      R_f[3,4] := -0.85727531;
      R_f[3,5] := 0.70266402;
      R_f[3,6] := -0.55573398;
      R_f[3,7] := 0.45469028;
      R_f[3,8] := -0.39782384;
      R_f[3,9] := 0.23143867;
      R_f[3,10] := -0.86177999;
      R_f[3,11] := 0.29983264;
      R_f[3,12] := 1.36218679;
      R_f[3,13] := 0.10939779;
      R_f[3,14] := -0.13315666;
      R_f[3,15] := -1.31117058;
      R_f[3,16] := 0.66998744;
      R_f[3,17] := 1.24320877;
      R_f[3,18] := -0.37031132;
      R_f[3,19] := -0.39300495;
      R_f[3,20] := -0.30342990;
      R_f[3,21] := -0.45216727;
      R_f[3,22] := -0.51143724;
      R_f[3,23] := 0.47799069;
      R_f[3,24] := -0.01827676;
      R_f[3,25] := 0.02519570;
      R_f[3,26] := 0.18636933;
      R_f[3,27] := -0.93594962;
      R_f[3,28] := 0.64644384;
      R_f[3,29] := -0.69783551;
      R_f[3,30] := -0.03558157;
      R_f[3,31] := 0.26994738;
      R_f[4,0] := -0.39344388;
      R_f[4,1] := 0.36222264;
      R_f[4,2] := -0.42310888;
      R_f[4,3] := 0.14989485;
      R_f[4,4] := -0.99088651;
      R_f[4,5] := 0.05782998;
      R_f[4,6] := 0.12812723;
      R_f[4,7] := -0.16467652;
      R_f[4,8] := -0.34736815;
      R_f[4,9] := 0.14911307;
      R_f[4,10] := 0.64495277;
      R_f[4,11] := 0.13966881;
      R_f[4,12] := 0.29640356;
      R_f[4,13] := 0.48785415;
      R_f[4,14] := -0.23574533;
      R_f[4,15] := 0.47339493;
      R_f[4,16] := -0.38768038;
      R_f[4,17] := 0.06993198;
      R_f[4,18] := 1.34699011;
      R_f[4,19] := -0.45494819;
      R_f[4,20] := -1.02421069;
      R_f[4,21] := 0.39080855;
      R_f[4,22] := -0.25200650;
      R_f[4,23] := 0.10465910;
      R_f[4,24] := 0.27367991;
      R_f[4,25] := 0.45886528;
      R_f[4,26] := 0.23802078;
      R_f[4,27] := -0.31698900;
      R_f[4,28] := 0.36807117;
      R_f[4,29] := -0.10262590;
      R_f[4,30] := -0.79831642;
      R_f[4,31] := 0.12268136;
      R_f[5,0] := 0.09268615;
      R_f[5,1] := 0.21935971;
      R_f[5,2] := -0.28605691;
      R_f[5,3] := -0.35209230;
      R_f[5,4] := 0.60323030;
      R_f[5,5] := -1.86963761;
      R_f[5,6] := 0.17267105;
      R_f[5,7] := 0.31667727;
      R_f[5,8] := 1.22614503;
      R_f[5,9] := -0.31814456;
      R_f[5,10] := 0.28639799;
      R_f[5,11] := 0.45808375;
      R_f[5,12] := 0.16454318;
      R_f[5,13] := -0.37628773;
      R_f[5,14] := 0.11079943;
      R_f[5,15] := 0.43248567;
      R_f[5,16] := 0.62867469;
      R_f[5,17] := -0.18534793;
      R_f[5,18] := -0.21310599;
      R_f[5,19] := -0.12530403;
      R_f[5,20] := -0.11672303;
      R_f[5,21] := -0.34058103;
      R_f[5,22] := 0.53213966;
      R_f[5,23] := -0.06069790;
      R_f[5,24] := 1.12480652;
      R_f[5,25] := -0.11877894;
      R_f[5,26] := 0.34038293;
      R_f[5,27] := 0.99329889;
      R_f[5,28] := 0.00048804;
      R_f[5,29] := -0.15688728;
      R_f[5,30] := 0.46641046;
      R_f[5,31] := 1.20925903;
      R_f[6,0] := -0.20363854;
      R_f[6,1] := -0.32236105;
      R_f[6,2] := -0.30276120;
      R_f[6,3] := -0.07836054;
      R_f[6,4] := 0.90966666;
      R_f[6,5] := 0.01400341;
      R_f[6,6] := 0.27368066;
      R_f[6,7] := 1.16410792;
      R_f[6,8] := 0.91342974;
      R_f[6,9] := -0.62499738;
      R_f[6,10] := 0.21230549;
      R_f[6,11] := 0.48843908;
      R_f[6,12] := -0.04002659;
      R_f[6,13] := -0.89160722;
      R_f[6,14] := 0.44720122;
      R_f[6,15] := -0.37033880;
      R_f[6,16] := 0.36007941;
      R_f[6,17] := 0.49022290;
      R_f[6,18] := -0.63365066;
      R_f[6,19] := -0.44222319;
      R_f[6,20] := 0.07470856;
      R_f[6,21] := -0.18424936;
      R_f[6,22] := -1.06331885;
      R_f[6,23] := 0.11231405;
      R_f[6,24] := 0.48846784;
      R_f[6,25] := 0.32240003;
      R_f[6,26] := -0.02514423;
      R_f[6,27] := 0.52824306;
      R_f[6,28] := 0.10916118;
      R_f[6,29] := 1.10423243;
      R_f[6,30] := 0.87132770;
      R_f[6,31] := -0.22497243;
      R_f[7,0] := 0.00290798;
      R_f[7,1] := 0.02380353;
      R_f[7,2] := -0.43460667;
      R_f[7,3] := -0.61469567;
      R_f[7,4] := 0.93173164;
      R_f[7,5] := -0.90107012;
      R_f[7,6] := 0.16509961;
      R_f[7,7] := 2.32758498;
      R_f[7,8] := -0.52484536;
      R_f[7,9] := 0.39195865;
      R_f[7,10] := -0.23609044;
      R_f[7,11] := 0.05608457;
      R_f[7,12] := -0.42776030;
      R_f[7,13] := -0.10564836;
      R_f[7,14] := -0.42611927;
      R_f[7,15] := -0.13254717;
      R_f[7,16] := 0.84613299;
      R_f[7,17] := -0.23140904;
      R_f[7,18] := 0.90073472;
      R_f[7,19] := -0.36597919;
      R_f[7,20] := 0.47446036;
      R_f[7,21] := -0.08705632;
      R_f[7,22] := -1.52176034;
      R_f[7,23] := 0.22270711;
      R_f[7,24] := -0.03422754;
      R_f[7,25] := 0.07659206;
      R_f[7,26] := 0.36599547;
      R_f[7,27] := -0.52767622;
      R_f[7,28] := -0.06631206;
      R_f[7,29] := -0.18978609;
      R_f[7,30] := 0.17292330;
      R_f[7,31] := 0.92969888;
      R_f[8,0] := -0.30634153;
      R_f[8,1] := -0.81952202;
      R_f[8,2] := -0.03526760;
      R_f[8,3] := -1.29526353;
      R_f[8,4] := 0.32094973;
      R_f[8,5] := -1.85603750;
      R_f[8,6] := 0.28356239;
      R_f[8,7] := 0.57538003;
      R_f[8,8] := -0.11039671;
      R_f[8,9] := -2.10963488;
      R_f[8,10] := -1.19219816;
      R_f[8,11] := -0.79363817;
      R_f[8,12] := 0.48992485;
      R_f[8,13] := 0.30308276;
      R_f[8,14] := 0.04908920;
      R_f[8,15] := 0.13945648;
      R_f[8,16] := -1.37335110;
      R_f[8,17] := 0.59385890;
      R_f[8,18] := -1.01455212;
      R_f[8,19] := -1.58437848;
      R_f[8,20] := -0.19760673;
      R_f[8,21] := -0.34158847;
      R_f[8,22] := 1.34096205;
      R_f[8,23] := 0.40719572;
      R_f[8,24] := -0.24326721;
      R_f[8,25] := -1.13661909;
      R_f[8,26] := -0.63606089;
      R_f[8,27] := 0.39769849;
      R_f[8,28] := -1.44548726;
      R_f[8,29] := 0.17782873;
      R_f[8,30] := -0.33304986;
      R_f[8,31] := -0.34794864;
      R_f[9,0] := -0.44309428;
      R_f[9,1] := -0.30440933;
      R_f[9,2] := 0.24199238;
      R_f[9,3] := 0.21034531;
      R_f[9,4] := -0.17321667;
      R_f[9,5] := -0.30677229;
      R_f[9,6] := -0.13734587;
      R_f[9,7] := 0.34537369;
      R_f[9,8] := -0.26872745;
      R_f[9,9] := 1.84128654;
      R_f[9,10] := 0.52121741;
      R_f[9,11] := 0.30513665;
      R_f[9,12] := -0.01998700;
      R_f[9,13] := -0.72075009;
      R_f[9,14] := -0.55062896;
      R_f[9,15] := -0.11161942;
      R_f[9,16] := 0.10928833;
      R_f[9,17] := 0.69333780;
      R_f[9,18] := -0.61185640;
      R_f[9,19] := -0.22928748;
      R_f[9,20] := 0.53006452;
      R_f[9,21] := 0.10420142;
      R_f[9,22] := -0.16613784;
      R_f[9,23] := 0.12584257;
      R_f[9,24] := 0.24575511;
      R_f[9,25] := 0.07394662;
      R_f[9,26] := 0.62375677;
      R_f[9,27] := 0.53293931;
      R_f[9,28] := 0.20416169;
      R_f[9,29] := -0.02031298;
      R_f[9,30] := -0.10528360;
      R_f[9,31] := 0.45511815;
      R_f[10,0] := 0.83232188;
      R_f[10,1] := -0.08258834;
      R_f[10,2] := -0.06935453;
      R_f[10,3] := 0.07768326;
      R_f[10,4] := 0.24524604;
      R_f[10,5] := -0.22525373;
      R_f[10,6] := 0.40935123;
      R_f[10,7] := -0.17911816;
      R_f[10,8] := -0.32271239;
      R_f[10,9] := -0.36832979;
      R_f[10,10] := -2.49958277;
      R_f[10,11] := -0.03748730;
      R_f[10,12] := -0.07992049;
      R_f[10,13] := 0.08578819;
      R_f[10,14] := -0.19220759;
      R_f[10,15] := 0.08966637;
      R_f[10,16] := -0.39432195;
      R_f[10,17] := 0.22714733;
      R_f[10,18] := -0.43346864;
      R_f[10,19] := -0.11305624;
      R_f[10,20] := 0.16338432;
      R_f[10,21] := -0.10953200;
      R_f[10,22] := -0.13001373;
      R_f[10,23] := 0.22707058;
      R_f[10,24] := 0.41991970;
      R_f[10,25] := 0.43455145;
      R_f[10,26] := 0.19583054;
      R_f[10,27] := 0.56395984;
      R_f[10,28] := -0.48473257;
      R_f[10,29] := 0.18865864;
      R_f[10,30] := 0.19654989;
      R_f[10,31] := 0.09913722;
      R_f[11,0] := 0.42754596;
      R_f[11,1] := 0.09423707;
      R_f[11,2] := -0.29017773;
      R_f[11,3] := -0.11189838;
      R_f[11,4] := -0.21009797;
      R_f[11,5] := -0.48191920;
      R_f[11,6] := 0.12651034;
      R_f[11,7] := 0.05790544;
      R_f[11,8] := -0.12319141;
      R_f[11,9] := 0.39675516;
      R_f[11,10] := -0.16217400;
      R_f[11,11] := 0.18192010;
      R_f[11,12] := 0.14949840;
      R_f[11,13] := -0.03762484;
      R_f[11,14] := -0.68928587;
      R_f[11,15] := 0.11334433;
      R_f[11,16] := -0.28812110;
      R_f[11,17] := 0.10144100;
      R_f[11,18] := -0.44992569;
      R_f[11,19] := -0.15579885;
      R_f[11,20] := -0.29591924;
      R_f[11,21] := -0.15366313;
      R_f[11,22] := -0.01909444;
      R_f[11,23] := 0.04565328;
      R_f[11,24] := -0.30796039;
      R_f[11,25] := -0.08308777;
      R_f[11,26] := 0.22044559;
      R_f[11,27] := 0.10441495;
      R_f[11,28] := 0.06342443;
      R_f[11,29] := -0.48254472;
      R_f[11,30] := 0.09183690;
      R_f[11,31] := -0.09384891;
      R_f[12,0] := 0.47012070;
      R_f[12,1] := -0.33459604;
      R_f[12,2] := -0.69821233;
      R_f[12,3] := 0.03733517;
      R_f[12,4] := 1.01428008;
      R_f[12,5] := -1.34689188;
      R_f[12,6] := 0.60434407;
      R_f[12,7] := 1.02553523;
      R_f[12,8] := 0.34444749;
      R_f[12,9] := -0.69957334;
      R_f[12,10] := 0.80366671;
      R_f[12,11] := 0.17610356;
      R_f[12,12] := 0.55641246;
      R_f[12,13] := -0.21217743;
      R_f[12,14] := -0.63918966;
      R_f[12,15] := -0.16232961;
      R_f[12,16] := 0.68742597;
      R_f[12,17] := 0.52715355;
      R_f[12,18] := 0.04790421;
      R_f[12,19] := -0.58621752;
      R_f[12,20] := 0.26796517;
      R_f[12,21] := -0.04791349;
      R_f[12,22] := -0.09341484;
      R_f[12,23] := 0.66781473;
      R_f[12,24] := 0.52626812;
      R_f[12,25] := 0.37837932;
      R_f[12,26] := 0.38251483;
      R_f[12,27] := 0.31467408;
      R_f[12,28] := -0.29517949;
      R_f[12,29] := -0.02343472;
      R_f[12,30] := 0.19953103;
      R_f[12,31] := 0.04299867;
      R_f[13,0] := 0.08943395;
      R_f[13,1] := -0.41928035;
      R_f[13,2] := -0.46420595;
      R_f[13,3] := -0.93849921;
      R_f[13,4] := 1.81882250;
      R_f[13,5] := -0.04638388;
      R_f[13,6] := -0.10525256;
      R_f[13,7] := -0.14901699;
      R_f[13,8] := 1.56855416;
      R_f[13,9] := -1.47332811;
      R_f[13,10] := 1.70304513;
      R_f[13,11] := 0.27727890;
      R_f[13,12] := 0.29618439;
      R_f[13,13] := 0.20549068;
      R_f[13,14] := 0.08464767;
      R_f[13,15] := -0.28658184;
      R_f[13,16] := 0.52141178;
      R_f[13,17] := -0.45672634;
      R_f[13,18] := -1.07117772;
      R_f[13,19] := -0.12635788;
      R_f[13,20] := -0.17076187;
      R_f[13,21] := -0.39133579;
      R_f[13,22] := -1.30128396;
      R_f[13,23] := -0.51295263;
      R_f[13,24] := 0.59420377;
      R_f[13,25] := -0.22949216;
      R_f[13,26] := -0.07507192;
      R_f[13,27] := 0.62209141;
      R_f[13,28] := -0.39097649;
      R_f[13,29] := 0.46184129;
      R_f[13,30] := 0.24478418;
      R_f[13,31] := 1.16894412;
      R_f[14,0] := 0.05281359;
      R_f[14,1] := -0.53310943;
      R_f[14,2] := -0.93560243;
      R_f[14,3] := 0.24883044;
      R_f[14,4] := -0.87425369;
      R_f[14,5] := 0.40351281;
      R_f[14,6] := -0.38772595;
      R_f[14,7] := 0.02093324;
      R_f[14,8] := -0.35284448;
      R_f[14,9] := -0.49149925;
      R_f[14,10] := 0.40103057;
      R_f[14,11] := -0.23631869;
      R_f[14,12] := -0.18181595;
      R_f[14,13] := 1.02885425;
      R_f[14,14] := 1.01850176;
      R_f[14,15] := 0.01374859;
      R_f[14,16] := 0.09904287;
      R_f[14,17] := 0.39969888;
      R_f[14,18] := 0.29445514;
      R_f[14,19] := -0.66422909;
      R_f[14,20] := 0.56930321;
      R_f[14,21] := 0.16506715;
      R_f[14,22] := -0.23321085;
      R_f[14,23] := 0.48102799;
      R_f[14,24] := -0.53297859;
      R_f[14,25] := 0.40016001;
      R_f[14,26] := -0.33044472;
      R_f[14,27] := 0.31068552;
      R_f[14,28] := 0.16014290;
      R_f[14,29] := 0.17083554;
      R_f[14,30] := 0.17105293;
      R_f[14,31] := 0.35666907;
      R_f[15,0] := 0.06514452;
      R_f[15,1] := -0.19740443;
      R_f[15,2] := 0.02617185;
      R_f[15,3] := 0.07652328;
      R_f[15,4] := 0.38803399;
      R_f[15,5] := -0.20535301;
      R_f[15,6] := -0.18448971;
      R_f[15,7] := -0.05007682;
      R_f[15,8] := -0.53877741;
      R_f[15,9] := 0.10129107;
      R_f[15,10] := 0.18535724;
      R_f[15,11] := 0.98206252;
      R_f[15,12] := 0.44447863;
      R_f[15,13] := -0.27786836;
      R_f[15,14] := -0.11058123;
      R_f[15,15] := 1.12241304;
      R_f[15,16] := 0.65275174;
      R_f[15,17] := -0.28105226;
      R_f[15,18] := -0.21099147;
      R_f[15,19] := 0.10379153;
      R_f[15,20] := -0.19425590;
      R_f[15,21] := -0.38361749;
      R_f[15,22] := -0.00013181;
      R_f[15,23] := -0.56550574;
      R_f[15,24] := 1.24397659;
      R_f[15,25] := 1.77377999;
      R_f[15,26] := 0.19124776;
      R_f[15,27] := 0.68570900;
      R_f[15,28] := -0.25024998;
      R_f[15,29] := -0.25333801;
      R_f[15,30] := 0.05722036;
      R_f[15,31] := 0.94418979;
      R_f[16,0] := 0.25488979;
      R_f[16,1] := -0.63715321;
      R_f[16,2] := 0.77243882;
      R_f[16,3] := 0.43674168;
      R_f[16,4] := 0.21674325;
      R_f[16,5] := -0.28702530;
      R_f[16,6] := 0.32552499;
      R_f[16,7] := -0.05745591;
      R_f[16,8] := 0.13758813;
      R_f[16,9] := -0.01359968;
      R_f[16,10] := -0.13954167;
      R_f[16,11] := 0.11212520;
      R_f[16,12] := 0.67787927;
      R_f[16,13] := 0.82328504;
      R_f[16,14] := -0.90781152;
      R_f[16,15] := -0.44112113;
      R_f[16,16] := 1.61208057;
      R_f[16,17] := -0.31707352;
      R_f[16,18] := 0.24660601;
      R_f[16,19] := -0.35153627;
      R_f[16,20] := -0.86473966;
      R_f[16,21] := -0.32204637;
      R_f[16,22] := 0.11319287;
      R_f[16,23] := 0.39265326;
      R_f[16,24] := -0.28525683;
      R_f[16,25] := -0.20465063;
      R_f[16,26] := -0.14012077;
      R_f[16,27] := -0.13221192;
      R_f[16,28] := 0.98584235;
      R_f[16,29] := 0.36052975;
      R_f[16,30] := -0.31423789;
      R_f[16,31] := 0.63994056;
      R_f[17,0] := 0.43413380;
      R_f[17,1] := -0.12179689;
      R_f[17,2] := -0.18103142;
      R_f[17,3] := -0.58753431;
      R_f[17,4] := 0.10463939;
      R_f[17,5] := -0.08838262;
      R_f[17,6] := 0.60563666;
      R_f[17,7] := 0.00878992;
      R_f[17,8] := -0.21168366;
      R_f[17,9] := 0.29472336;
      R_f[17,10] := 0.22692770;
      R_f[17,11] := 0.27634826;
      R_f[17,12] := -0.16206916;
      R_f[17,13] := -0.25042766;
      R_f[17,14] := -0.24090815;
      R_f[17,15] := 0.28610602;
      R_f[17,16] := -0.55426306;
      R_f[17,17] := 1.41948617;
      R_f[17,18] := 0.40432185;
      R_f[17,19] := 0.47929171;
      R_f[17,20] := -0.07214013;
      R_f[17,21] := 0.10474437;
      R_f[17,22] := 0.05560365;
      R_f[17,23] := 0.29282579;
      R_f[17,24] := -0.02698746;
      R_f[17,25] := 0.45795625;
      R_f[17,26] := 0.45755112;
      R_f[17,27] := -0.19397356;
      R_f[17,28] := -0.22833887;
      R_f[17,29] := -0.40156868;
      R_f[17,30] := -0.06691723;
      R_f[17,31] := -0.16601346;
      R_f[18,0] := 0.21388659;
      R_f[18,1] := -0.21044491;
      R_f[18,2] := -0.18511969;
      R_f[18,3] := 0.12251608;
      R_f[18,4] := -0.82450879;
      R_f[18,5] := -0.50903809;
      R_f[18,6] := -0.44293392;
      R_f[18,7] := 0.31674486;
      R_f[18,8] := -0.11843041;
      R_f[18,9] := -0.19616166;
      R_f[18,10] := 0.17610525;
      R_f[18,11] := 0.51645488;
      R_f[18,12] := 0.46033934;
      R_f[18,13] := 0.35017881;
      R_f[18,14] := 0.49660042;
      R_f[18,15] := 0.02593680;
      R_f[18,16] := 0.25847656;
      R_f[18,17] := -0.18605545;
      R_f[18,18] := 1.64782512;
      R_f[18,19] := -0.23618795;
      R_f[18,20] := -0.00984277;
      R_f[18,21] := -0.22337262;
      R_f[18,22] := 0.01971689;
      R_f[18,23] := -0.08102468;
      R_f[18,24] := -0.63402730;
      R_f[18,25] := -0.07497400;
      R_f[18,26] := 0.15719052;
      R_f[18,27] := -0.07695547;
      R_f[18,28] := -0.27590719;
      R_f[18,29] := 0.31225580;
      R_f[18,30] := 0.20215666;
      R_f[18,31] := -0.08998311;
      R_f[19,0] := 0.46975327;
      R_f[19,1] := 0.17221756;
      R_f[19,2] := 0.17129607;
      R_f[19,3] := 0.05666168;
      R_f[19,4] := 0.14368458;
      R_f[19,5] := -0.54253471;
      R_f[19,6] := 0.40939260;
      R_f[19,7] := 0.05611381;
      R_f[19,8] := -0.78961420;
      R_f[19,9] := 0.35195425;
      R_f[19,10] := 0.16296588;
      R_f[19,11] := 0.54626679;
      R_f[19,12] := -0.08277176;
      R_f[19,13] := -0.22074869;
      R_f[19,14] := -0.65805823;
      R_f[19,15] := -0.05598476;
      R_f[19,16] := -0.04306423;
      R_f[19,17] := -0.32691059;
      R_f[19,18] := -0.33659294;
      R_f[19,19] := -1.07530594;
      R_f[19,20] := 0.17525475;
      R_f[19,21] := -0.07675232;
      R_f[19,22] := 0.10386194;
      R_f[19,23] := 0.19622359;
      R_f[19,24] := 0.17771964;
      R_f[19,25] := -0.01513422;
      R_f[19,26] := 0.36328980;
      R_f[19,27] := 0.06220879;
      R_f[19,28] := -0.39328694;
      R_f[19,29] := 0.33954379;
      R_f[19,30] := 0.05713883;
      R_f[19,31] := -0.33563131;
      R_f[20,0] := 0.18057881;
      R_f[20,1] := -0.24642186;
      R_f[20,2] := -0.24286529;
      R_f[20,3] := -0.67373210;
      R_f[20,4] := 0.90808105;
      R_f[20,5] := -1.08204496;
      R_f[20,6] := -0.78024036;
      R_f[20,7] := 1.16503656;
      R_f[20,8] := 0.43974155;
      R_f[20,9] := -1.03952718;
      R_f[20,10] := -0.28429365;
      R_f[20,11] := -0.25702575;
      R_f[20,12] := -0.15614110;
      R_f[20,13] := -0.04867256;
      R_f[20,14] := 1.24517381;
      R_f[20,15] := -0.50706828;
      R_f[20,16] := -0.20075536;
      R_f[20,17] := 0.10849988;
      R_f[20,18] := 0.75873327;
      R_f[20,19] := -0.02426600;
      R_f[20,20] := -1.02889967;
      R_f[20,21] := -0.49422511;
      R_f[20,22] := 0.76041186;
      R_f[20,23] := -0.04359674;
      R_f[20,24] := -0.15679558;
      R_f[20,25] := -0.14447898;
      R_f[20,26] := -0.46510464;
      R_f[20,27] := 1.35692060;
      R_f[20,28] := -0.93135232;
      R_f[20,29] := 0.77650243;
      R_f[20,30] := -0.63533545;
      R_f[20,31] := 0.93425041;
      R_f[21,0] := 0.41408271;
      R_f[21,1] := -0.37474987;
      R_f[21,2] := 0.06901271;
      R_f[21,3] := 0.05882899;
      R_f[21,4] := 1.50155163;
      R_f[21,5] := -0.68119925;
      R_f[21,6] := -0.99283367;
      R_f[21,7] := -0.16499096;
      R_f[21,8] := -0.39376357;
      R_f[21,9] := -1.37646723;
      R_f[21,10] := 0.64534718;
      R_f[21,11] := 0.08503322;
      R_f[21,12] := 0.22116974;
      R_f[21,13] := -0.18298884;
      R_f[21,14] := -0.00657548;
      R_f[21,15] := -0.18632370;
      R_f[21,16] := -0.26151741;
      R_f[21,17] := -0.03215327;
      R_f[21,18] := -1.32762277;
      R_f[21,19] := 0.35820487;
      R_f[21,20] := -0.43136457;
      R_f[21,21] := 0.08935426;
      R_f[21,22] := 0.23742658;
      R_f[21,23] := 0.30326349;
      R_f[21,24] := 1.07324779;
      R_f[21,25] := -0.18277077;
      R_f[21,26] := -0.06333762;
      R_f[21,27] := -0.08517780;
      R_f[21,28] := -1.28671491;
      R_f[21,29] := -0.49619201;
      R_f[21,30] := -0.18604164;
      R_f[21,31] := 1.17694867;
      R_f[22,0] := -0.35642302;
      R_f[22,1] := -0.07537675;
      R_f[22,2] := -0.11212978;
      R_f[22,3] := 0.91988707;
      R_f[22,4] := 0.29476365;
      R_f[22,5] := -0.08478891;
      R_f[22,6] := 0.06471095;
      R_f[22,7] := 1.18266797;
      R_f[22,8] := 0.17392084;
      R_f[22,9] := -0.08943880;
      R_f[22,10] := 0.23702587;
      R_f[22,11] := -0.43714434;
      R_f[22,12] := 0.07848407;
      R_f[22,13] := -0.14684126;
      R_f[22,14] := 0.02883088;
      R_f[22,15] := -0.60347939;
      R_f[22,16] := 0.02053990;
      R_f[22,17] := 0.93891013;
      R_f[22,18] := 0.25982085;
      R_f[22,19] := 0.18691589;
      R_f[22,20] := -0.16190472;
      R_f[22,21] := -0.56379879;
      R_f[22,22] := 1.18819308;
      R_f[22,23] := 0.14459842;
      R_f[22,24] := 0.38293535;
      R_f[22,25] := -0.46581766;
      R_f[22,26] := 0.53433573;
      R_f[22,27] := 0.16328283;
      R_f[22,28] := 0.04261781;
      R_f[22,29] := -0.32524684;
      R_f[22,30] := 0.08497128;
      R_f[22,31] := 0.73156911;
      R_f[23,0] := -0.04014154;
      R_f[23,1] := -0.21957491;
      R_f[23,2] := -0.47944790;
      R_f[23,3] := -0.18949568;
      R_f[23,4] := 0.20813392;
      R_f[23,5] := -1.26923680;
      R_f[23,6] := -0.43531770;
      R_f[23,7] := 0.03713821;
      R_f[23,8] := 0.59817761;
      R_f[23,9] := -0.59432054;
      R_f[23,10] := 0.37402180;
      R_f[23,11] := -0.15723693;
      R_f[23,12] := 0.19139190;
      R_f[23,13] := -0.80456918;
      R_f[23,14] := -0.05263249;
      R_f[23,15] := -0.29430014;
      R_f[23,16] := 0.26987091;
      R_f[23,17] := 0.34275058;
      R_f[23,18] := 0.44585946;
      R_f[23,19] := -0.86910695;
      R_f[23,20] := -1.37904131;
      R_f[23,21] := 0.03121136;
      R_f[23,22] := 0.20768139;
      R_f[23,23] := 0.96365720;
      R_f[23,24] := 1.29164517;
      R_f[23,25] := 0.27564162;
      R_f[23,26] := 0.19493468;
      R_f[23,27] := 0.25765347;
      R_f[23,28] := -0.75100589;
      R_f[23,29] := 0.41528577;
      R_f[23,30] := 1.09287107;
      R_f[23,31] := 0.43580219;
      R_f[24,0] := 0.10901141;
      R_f[24,1] := -0.00615504;
      R_f[24,2] := -0.42680290;
      R_f[24,3] := -0.48820597;
      R_f[24,4] := 1.09372568;
      R_f[24,5] := -0.64686328;
      R_f[24,6] := 0.10192143;
      R_f[24,7] := 0.28666073;
      R_f[24,8] := 0.64033169;
      R_f[24,9] := -1.23651469;
      R_f[24,10] := 0.14855224;
      R_f[24,11] := -0.15615174;
      R_f[24,12] := -0.25834996;
      R_f[24,13] := -0.13889249;
      R_f[24,14] := 0.62434721;
      R_f[24,15] := -0.46040115;
      R_f[24,16] := -0.01414216;
      R_f[24,17] := -0.28662860;
      R_f[24,18] := -0.24730733;
      R_f[24,19] := -0.03740590;
      R_f[24,20] := 0.03079495;
      R_f[24,21] := -1.07491624;
      R_f[24,22] := -0.32715502;
      R_f[24,23] := 0.03199894;
      R_f[24,24] := -0.06877741;
      R_f[24,25] := 0.12599984;
      R_f[24,26] := -0.46782377;
      R_f[24,27] := 0.64110184;
      R_f[24,28] := 0.04548985;
      R_f[24,29] := 0.05152436;
      R_f[24,30] := 0.15953350;
      R_f[24,31] := 0.43480337;
      R_f[25,0] := 1.16320372;
      R_f[25,1] := 0.06548461;
      R_f[25,2] := 0.28802359;
      R_f[25,3] := 0.55442971;
      R_f[25,4] := 0.25373462;
      R_f[25,5] := -0.37025258;
      R_f[25,6] := -0.48865169;
      R_f[25,7] := 0.16444007;
      R_f[25,8] := 0.16262302;
      R_f[25,9] := -0.28667378;
      R_f[25,10] := -1.04200613;
      R_f[25,11] := -0.24463102;
      R_f[25,12] := 0.26678899;
      R_f[25,13] := -0.35289085;
      R_f[25,14] := 0.45832568;
      R_f[25,15] := 0.08287992;
      R_f[25,16] := -0.90763897;
      R_f[25,17] := 1.16429114;
      R_f[25,18] := -0.51552850;
      R_f[25,19] := -0.00712482;
      R_f[25,20] := 0.10827811;
      R_f[25,21] := 0.30554232;
      R_f[25,22] := -0.13470046;
      R_f[25,23] := -0.05728173;
      R_f[25,24] := 0.25545090;
      R_f[25,25] := 1.25365567;
      R_f[25,26] := 0.49803498;
      R_f[25,27] := 1.85552025;
      R_f[25,28] := -1.15144587;
      R_f[25,29] := 0.07574563;
      R_f[25,30] := 1.53851593;
      R_f[25,31] := -0.06473381;
      R_f[26,0] := 0.59528756;
      R_f[26,1] := -0.18308367;
      R_f[26,2] := 0.34858477;
      R_f[26,3] := -0.04807191;
      R_f[26,4] := 1.62759721;
      R_f[26,5] := -1.32408214;
      R_f[26,6] := -0.86638910;
      R_f[26,7] := 0.98388058;
      R_f[26,8] := 0.84169364;
      R_f[26,9] := -0.06820829;
      R_f[26,10] := 0.92988855;
      R_f[26,11] := -0.03296947;
      R_f[26,12] := 1.13297725;
      R_f[26,13] := -0.57467204;
      R_f[26,14] := 0.52196753;
      R_f[26,15] := 0.43573204;
      R_f[26,16] := 1.07805049;
      R_f[26,17] := 0.23477279;
      R_f[26,18] := -0.39657351;
      R_f[26,19] := 0.55390966;
      R_f[26,20] := -0.07512384;
      R_f[26,21] := -0.93572176;
      R_f[26,22] := 0.54867393;
      R_f[26,23] := -0.29351887;
      R_f[26,24] := 0.28448883;
      R_f[26,25] := 0.72720629;
      R_f[26,26] := 1.01896834;
      R_f[26,27] := -0.14029346;
      R_f[26,28] := -0.65743059;
      R_f[26,29] := -0.32555410;
      R_f[26,30] := 1.61288857;
      R_f[26,31] := 0.18683940;
      R_f[27,0] := -0.80839366;
      R_f[27,1] := -0.49256265;
      R_f[27,2] := -0.46127644;
      R_f[27,3] := -0.26435462;
      R_f[27,4] := 0.45098844;
      R_f[27,5] := -0.50330544;
      R_f[27,6] := -0.20470831;
      R_f[27,7] := 0.94890404;
      R_f[27,8] := -0.01666292;
      R_f[27,9] := -0.45548967;
      R_f[27,10] := 0.61688972;
      R_f[27,11] := 0.71183705;
      R_f[27,12] := -0.24694404;
      R_f[27,13] := 0.12021586;
      R_f[27,14] := -0.04486329;
      R_f[27,15] := -0.39616454;
      R_f[27,16] := 0.51417869;
      R_f[27,17] := -0.39478543;
      R_f[27,18] := 0.25215191;
      R_f[27,19] := -0.16793472;
      R_f[27,20] := -0.11071328;
      R_f[27,21] := 0.02187885;
      R_f[27,22] := 0.26461548;
      R_f[27,23] := -0.31467691;
      R_f[27,24] := 0.06920367;
      R_f[27,25] := -0.56788224;
      R_f[27,26] := -0.61690986;
      R_f[27,27] := -0.68749779;
      R_f[27,28] := -1.40037727;
      R_f[27,29] := 0.65967739;
      R_f[27,30] := -1.72095454;
      R_f[27,31] := 1.51459014;
      R_f[28,0] := 0.53473991;
      R_f[28,1] := 0.12026238;
      R_f[28,2] := -0.44487497;
      R_f[28,3] := 0.11609860;
      R_f[28,4] := -0.09671389;
      R_f[28,5] := 0.03561250;
      R_f[28,6] := -0.00043401;
      R_f[28,7] := -0.22344112;
      R_f[28,8] := -0.74334919;
      R_f[28,9] := 0.22675149;
      R_f[28,10] := -0.02913556;
      R_f[28,11] := 0.67491484;
      R_f[28,12] := -0.26046002;
      R_f[28,13] := 0.23686388;
      R_f[28,14] := -0.16231716;
      R_f[28,15] := 0.22020151;
      R_f[28,16] := 0.22111253;
      R_f[28,17] := -0.28245488;
      R_f[28,18] := 0.43832338;
      R_f[28,19] := 0.56766087;
      R_f[28,20] := 0.12882017;
      R_f[28,21] := 0.34402338;
      R_f[28,22] := -0.13627987;
      R_f[28,23] := 0.05657256;
      R_f[28,24] := -0.43770042;
      R_f[28,25] := 0.52974325;
      R_f[28,26] := 0.55016619;
      R_f[28,27] := 0.32488731;
      R_f[28,28] := 0.31555337;
      R_f[28,29] := -0.32505563;
      R_f[28,30] := -0.54369146;
      R_f[28,31] := -0.21397509;
      R_f[29,0] := 0.74640977;
      R_f[29,1] := -0.51247251;
      R_f[29,2] := -0.71097630;
      R_f[29,3] := -0.90446025;
      R_f[29,4] := 0.44504565;
      R_f[29,5] := -0.89021724;
      R_f[29,6] := 0.81150109;
      R_f[29,7] := 0.45580223;
      R_f[29,8] := 0.48597828;
      R_f[29,9] := -0.12246494;
      R_f[29,10] := 0.75742763;
      R_f[29,11] := 0.15665157;
      R_f[29,12] := 0.99491531;
      R_f[29,13] := -0.29243794;
      R_f[29,14] := -0.63920891;
      R_f[29,15] := -0.07434531;
      R_f[29,16] := 0.64870352;
      R_f[29,17] := 0.26328391;
      R_f[29,18] := -0.64544326;
      R_f[29,19] := 0.55969763;
      R_f[29,20] := -1.23505473;
      R_f[29,21] := -1.08088791;
      R_f[29,22] := 0.23190728;
      R_f[29,23] := 0.33156013;
      R_f[29,24] := 1.42430663;
      R_f[29,25] := 0.83351737;
      R_f[29,26] := 0.95834678;
      R_f[29,27] := 0.52043319;
      R_f[29,28] := -0.28924993;
      R_f[29,29] := -1.70719016;
      R_f[29,30] := 0.81097376;
      R_f[29,31] := 1.26607156;
      R_f[30,0] := 0.18132812;
      R_f[30,1] := -0.38076901;
      R_f[30,2] := -0.33011848;
      R_f[30,3] := 0.09190890;
      R_f[30,4] := 0.40049037;
      R_f[30,5] := -0.56039268;
      R_f[30,6] := 0.04094384;
      R_f[30,7] := 0.67939031;
      R_f[30,8] := -0.18653642;
      R_f[30,9] := -0.43633384;
      R_f[30,10] := 0.27230042;
      R_f[30,11] := 0.39263970;
      R_f[30,12] := 0.33082095;
      R_f[30,13] := -0.07204608;
      R_f[30,14] := -0.16458063;
      R_f[30,15] := 0.11422759;
      R_f[30,16] := -0.02973648;
      R_f[30,17] := -0.61857194;
      R_f[30,18] := 0.20339146;
      R_f[30,19] := -0.12102985;
      R_f[30,20] := -0.23646855;
      R_f[30,21] := 0.16910897;
      R_f[30,22] := 0.05366793;
      R_f[30,23] := 0.17361535;
      R_f[30,24] := 0.07103206;
      R_f[30,25] := -0.02880308;
      R_f[30,26] := 0.10739103;
      R_f[30,27] := -0.29030880;
      R_f[30,28] := -0.03621915;
      R_f[30,29] := 0.09102457;
      R_f[30,30] := -1.78858960;
      R_f[30,31] := 0.76714230;
      R_f[31,0] := 0.52647686;
      R_f[31,1] := -0.90124124;
      R_f[31,2] := -0.03594093;
      R_f[31,3] := -0.14132296;
      R_f[31,4] := 0.02861782;
      R_f[31,5] := -0.32323492;
      R_f[31,6] := 0.83903587;
      R_f[31,7] := 0.13043062;
      R_f[31,8] := 0.03886109;
      R_f[31,9] := -1.15255368;
      R_f[31,10] := 0.28511661;
      R_f[31,11] := 0.14256424;
      R_f[31,12] := 0.14117993;
      R_f[31,13] := -0.76906091;
      R_f[31,14] := 0.29417679;
      R_f[31,15] := -0.36273482;
      R_f[31,16] := 0.45405060;
      R_f[31,17] := 0.05709918;
      R_f[31,18] := -0.90280342;
      R_f[31,19] := -0.48238260;
      R_f[31,20] := 0.38758871;
      R_f[31,21] := -0.09756728;
      R_f[31,22] := -0.48481289;
      R_f[31,23] := 0.10114307;
      R_f[31,24] := 0.44602498;
      R_f[31,25] := 0.42367566;
      R_f[31,26] := 0.35134542;
      R_f[31,27] := 2.05784130;
      R_f[31,28] := 0.03545408;
      R_f[31,29] := -0.16603291;
      R_f[31,30] := 0.86331582;
      R_f[31,31] := 2.59947228;
      R_g[0,0] := -3.21544218;
      R_g[0,1] := 0.04580142;
      R_g[0,2] := 0.06932437;
      R_g[0,3] := -0.15209895;
      R_g[0,4] := -0.09220740;
      R_g[0,5] := -0.07005115;
      R_g[0,6] := -0.24692968;
      R_g[0,7] := -0.08400031;
      R_g[0,8] := 0.17623347;
      R_g[0,9] := 0.00386813;
      R_g[0,10] := 0.06843853;
      R_g[0,11] := 0.21401274;
      R_g[0,12] := -0.15987185;
      R_g[0,13] := 0.24538136;
      R_g[0,14] := -0.18053962;
      R_g[0,15] := 0.34869576;
      R_g[0,16] := 0.01967172;
      R_g[0,17] := 0.15144458;
      R_g[0,18] := 0.11171592;
      R_g[0,19] := -0.15803322;
      R_g[0,20] := -0.16891836;
      R_g[0,21] := -0.05628303;
      R_g[0,22] := -0.31057128;
      R_g[0,23] := -0.08424718;
      R_g[0,24] := -0.00991914;
      R_g[0,25] := 0.02045443;
      R_g[0,26] := -0.58750242;
      R_g[0,27] := -0.19864596;
      R_g[0,28] := 0.02947442;
      R_g[0,29] := -0.11766856;
      R_g[0,30] := 0.03604466;
      R_g[0,31] := 0.00360318;
      R_g[1,0] := -0.31844607;
      R_g[1,1] := -6.12028122;
      R_g[1,2] := -0.26272821;
      R_g[1,3] := -0.13002822;
      R_g[1,4] := -0.32366905;
      R_g[1,5] := -0.18344826;
      R_g[1,6] := 0.68305010;
      R_g[1,7] := -0.09005546;
      R_g[1,8] := 0.54662579;
      R_g[1,9] := 0.13805637;
      R_g[1,10] := 0.02323161;
      R_g[1,11] := -0.34067392;
      R_g[1,12] := -0.17073138;
      R_g[1,13] := 0.39132595;
      R_g[1,14] := -0.18808186;
      R_g[1,15] := -0.26003635;
      R_g[1,16] := -0.19648901;
      R_g[1,17] := 0.16843174;
      R_g[1,18] := 0.15324172;
      R_g[1,19] := 0.45543799;
      R_g[1,20] := -0.65539354;
      R_g[1,21] := 0.56102079;
      R_g[1,22] := 0.13624945;
      R_g[1,23] := 0.21319284;
      R_g[1,24] := -0.25470603;
      R_g[1,25] := 0.26430780;
      R_g[1,26] := 0.27211225;
      R_g[1,27] := 0.04482314;
      R_g[1,28] := 0.01593675;
      R_g[1,29] := -0.23828241;
      R_g[1,30] := -0.16030560;
      R_g[1,31] := -0.15435591;
      R_g[2,0] := 0.54044676;
      R_g[2,1] := 0.45466635;
      R_g[2,2] := -4.12347174;
      R_g[2,3] := 0.41999578;
      R_g[2,4] := 0.72307265;
      R_g[2,5] := -0.14744292;
      R_g[2,6] := 0.76321173;
      R_g[2,7] := -0.18524313;
      R_g[2,8] := 0.11785751;
      R_g[2,9] := -0.17083235;
      R_g[2,10] := -0.22937453;
      R_g[2,11] := 0.00189192;
      R_g[2,12] := -0.26274452;
      R_g[2,13] := -0.87501872;
      R_g[2,14] := -0.28829265;
      R_g[2,15] := -0.56726843;
      R_g[2,16] := 0.72544920;
      R_g[2,17] := 0.59341317;
      R_g[2,18] := -0.24143113;
      R_g[2,19] := 0.12870285;
      R_g[2,20] := 0.14126211;
      R_g[2,21] := -0.39131889;
      R_g[2,22] := 0.25232065;
      R_g[2,23] := -0.38939855;
      R_g[2,24] := 0.55910432;
      R_g[2,25] := -0.29941782;
      R_g[2,26] := -0.28899693;
      R_g[2,27] := -0.10321512;
      R_g[2,28] := -0.40149158;
      R_g[2,29] := -0.11851617;
      R_g[2,30] := -0.12619454;
      R_g[2,31] := -0.27980283;
      R_g[3,0] := -0.53001744;
      R_g[3,1] := -0.11381795;
      R_g[3,2] := 0.11633322;
      R_g[3,3] := -0.43659294;
      R_g[3,4] := -0.60524720;
      R_g[3,5] := 0.05234856;
      R_g[3,6] := -0.46642643;
      R_g[3,7] := 0.27130726;
      R_g[3,8] := 0.09782532;
      R_g[3,9] := 0.38945866;
      R_g[3,10] := 0.14257543;
      R_g[3,11] := 0.58669364;
      R_g[3,12] := 0.55071652;
      R_g[3,13] := 0.51357007;
      R_g[3,14] := -0.08788987;
      R_g[3,15] := 0.94994968;
      R_g[3,16] := -0.44708440;
      R_g[3,17] := 0.02437577;
      R_g[3,18] := 0.58858347;
      R_g[3,19] := -0.45520020;
      R_g[3,20] := -0.09173007;
      R_g[3,21] := 0.72423649;
      R_g[3,22] := -0.38213339;
      R_g[3,23] := 0.50569993;
      R_g[3,24] := -0.41009858;
      R_g[3,25] := 0.38796568;
      R_g[3,26] := -0.68482327;
      R_g[3,27] := -0.01562345;
      R_g[3,28] := 0.03469054;
      R_g[3,29] := 0.34822434;
      R_g[3,30] := -0.32064009;
      R_g[3,31] := -0.42251477;
      R_g[4,0] := -0.02385795;
      R_g[4,1] := 0.39379948;
      R_g[4,2] := 0.10996556;
      R_g[4,3] := -0.30819508;
      R_g[4,4] := 0.00654567;
      R_g[4,5] := 0.20766497;
      R_g[4,6] := 0.13965006;
      R_g[4,7] := 0.04763399;
      R_g[4,8] := -0.12334181;
      R_g[4,9] := -0.29001412;
      R_g[4,10] := 0.27730298;
      R_g[4,11] := -0.03456333;
      R_g[4,12] := 0.27051720;
      R_g[4,13] := -1.29572177;
      R_g[4,14] := 0.32791910;
      R_g[4,15] := -0.26211676;
      R_g[4,16] := -0.34868079;
      R_g[4,17] := -0.59147680;
      R_g[4,18] := 0.38750806;
      R_g[4,19] := 0.30694690;
      R_g[4,20] := -0.06771316;
      R_g[4,21] := 0.07994391;
      R_g[4,22] := -0.20993046;
      R_g[4,23] := 0.01419108;
      R_g[4,24] := 1.40602803;
      R_g[4,25] := -0.26541275;
      R_g[4,26] := -0.25228849;
      R_g[4,27] := 0.49503145;
      R_g[4,28] := 0.01375614;
      R_g[4,29] := -0.36419708;
      R_g[4,30] := -0.03669171;
      R_g[4,31] := 1.10761940;
      R_g[5,0] := -0.06672658;
      R_g[5,1] := 0.04556764;
      R_g[5,2] := -0.34957722;
      R_g[5,3] := 0.09752260;
      R_g[5,4] := -0.26705503;
      R_g[5,5] := -4.08511257;
      R_g[5,6] := 0.36573645;
      R_g[5,7] := 0.02826878;
      R_g[5,8] := -0.27328387;
      R_g[5,9] := -0.18392695;
      R_g[5,10] := -0.06489211;
      R_g[5,11] := -0.17845686;
      R_g[5,12] := 0.02167919;
      R_g[5,13] := -0.11682998;
      R_g[5,14] := -0.07696812;
      R_g[5,15] := -0.01392019;
      R_g[5,16] := 0.48726702;
      R_g[5,17] := 0.01458673;
      R_g[5,18] := 0.74653000;
      R_g[5,19] := -0.70791829;
      R_g[5,20] := -0.20737875;
      R_g[5,21] := 0.33243728;
      R_g[5,22] := 0.03939781;
      R_g[5,23] := 0.11626533;
      R_g[5,24] := -0.13828859;
      R_g[5,25] := 0.04565351;
      R_g[5,26] := 0.20426168;
      R_g[5,27] := 0.25344858;
      R_g[5,28] := 0.07790031;
      R_g[5,29] := -0.33917236;
      R_g[5,30] := 0.20142451;
      R_g[5,31] := -0.03987967;
      R_g[6,0] := 0.34297273;
      R_g[6,1] := 0.14082512;
      R_g[6,2] := -0.00792844;
      R_g[6,3] := 0.46256095;
      R_g[6,4] := 0.15239693;
      R_g[6,5] := -0.36170921;
      R_g[6,6] := -4.22906876;
      R_g[6,7] := 0.26568046;
      R_g[6,8] := 0.11281063;
      R_g[6,9] := -0.54930890;
      R_g[6,10] := -0.38224915;
      R_g[6,11] := 0.21145333;
      R_g[6,12] := 0.15898399;
      R_g[6,13] := 0.56838512;
      R_g[6,14] := 0.26312956;
      R_g[6,15] := -0.45246279;
      R_g[6,16] := 0.45148721;
      R_g[6,17] := 0.18431610;
      R_g[6,18] := -0.27582157;
      R_g[6,19] := 0.17563862;
      R_g[6,20] := -0.07097334;
      R_g[6,21] := 0.15246704;
      R_g[6,22] := 0.05121115;
      R_g[6,23] := -0.15158200;
      R_g[6,24] := -0.01810670;
      R_g[6,25] := -0.12762244;
      R_g[6,26] := -0.77893329;
      R_g[6,27] := -0.29004732;
      R_g[6,28] := -0.19388825;
      R_g[6,29] := -0.31783766;
      R_g[6,30] := -0.26640892;
      R_g[6,31] := 0.22308391;
      R_g[7,0] := -0.26773775;
      R_g[7,1] := 0.25460386;
      R_g[7,2] := 0.00816728;
      R_g[7,3] := -0.20814449;
      R_g[7,4] := -0.12277725;
      R_g[7,5] := -0.12499115;
      R_g[7,6] := -0.06594294;
      R_g[7,7] := -4.17999268;
      R_g[7,8] := 0.25158358;
      R_g[7,9] := 0.38836476;
      R_g[7,10] := 0.12598813;
      R_g[7,11] := -0.03031898;
      R_g[7,12] := -0.67921215;
      R_g[7,13] := 0.16266112;
      R_g[7,14] := -0.25174144;
      R_g[7,15] := 0.33827740;
      R_g[7,16] := -0.28344563;
      R_g[7,17] := 0.38798764;
      R_g[7,18] := 0.28595367;
      R_g[7,19] := 0.02082766;
      R_g[7,20] := -0.42146638;
      R_g[7,21] := -0.23499288;
      R_g[7,22] := -0.01005266;
      R_g[7,23] := -0.06581271;
      R_g[7,24] := 0.08085475;
      R_g[7,25] := 0.06523639;
      R_g[7,26] := -0.14278226;
      R_g[7,27] := -0.05057906;
      R_g[7,28] := -0.17726235;
      R_g[7,29] := -0.15383634;
      R_g[7,30] := -0.07735643;
      R_g[7,31] := -0.52492666;
      R_g[8,0] := -0.05682376;
      R_g[8,1] := 0.08511543;
      R_g[8,2] := -0.11766159;
      R_g[8,3] := -0.10838570;
      R_g[8,4] := 0.00487707;
      R_g[8,5] := 0.14100854;
      R_g[8,6] := 0.34960595;
      R_g[8,7] := -0.48418933;
      R_g[8,8] := -3.81799150;
      R_g[8,9] := 0.63066083;
      R_g[8,10] := 0.84131134;
      R_g[8,11] := 0.11601801;
      R_g[8,12] := -0.44023189;
      R_g[8,13] := -0.08075541;
      R_g[8,14] := -0.23601621;
      R_g[8,15] := 0.16050224;
      R_g[8,16] := 0.11950148;
      R_g[8,17] := 0.87579739;
      R_g[8,18] := 0.89856052;
      R_g[8,19] := 1.38507712;
      R_g[8,20] := 0.29738313;
      R_g[8,21] := -0.01374565;
      R_g[8,22] := -0.33392283;
      R_g[8,23] := 0.01949951;
      R_g[8,24] := -0.09455296;
      R_g[8,25] := 0.24886662;
      R_g[8,26] := 0.05108426;
      R_g[8,27] := -0.13569650;
      R_g[8,28] := -0.14587976;
      R_g[8,29] := 0.29113290;
      R_g[8,30] := -0.01038904;
      R_g[8,31] := 0.19652341;
      R_g[9,0] := 0.38026151;
      R_g[9,1] := 0.14169994;
      R_g[9,2] := 0.37200066;
      R_g[9,3] := 0.15880315;
      R_g[9,4] := 0.10081743;
      R_g[9,5] := 0.13654961;
      R_g[9,6] := 1.48897541;
      R_g[9,7] := -0.10697847;
      R_g[9,8] := 0.39174217;
      R_g[9,9] := -1.73796725;
      R_g[9,10] := 0.19905937;
      R_g[9,11] := -0.08040750;
      R_g[9,12] := -0.53451943;
      R_g[9,13] := 0.30285180;
      R_g[9,14] := -0.34968182;
      R_g[9,15] := 0.19448446;
      R_g[9,16] := 0.52780533;
      R_g[9,17] := 0.89234567;
      R_g[9,18] := -0.13963117;
      R_g[9,19] := -0.33441579;
      R_g[9,20] := -0.37530658;
      R_g[9,21] := 0.16917522;
      R_g[9,22] := -0.43314484;
      R_g[9,23] := 0.37773979;
      R_g[9,24] := -0.26563615;
      R_g[9,25] := 0.27597877;
      R_g[9,26] := -0.59992433;
      R_g[9,27] := -1.16615653;
      R_g[9,28] := 0.34234476;
      R_g[9,29] := -0.21711856;
      R_g[9,30] := -0.15369894;
      R_g[9,31] := 0.00771751;
      R_g[10,0] := 0.06583999;
      R_g[10,1] := 0.08891983;
      R_g[10,2] := -0.57995307;
      R_g[10,3] := -0.03708947;
      R_g[10,4] := 0.65756792;
      R_g[10,5] := -0.66560614;
      R_g[10,6] := -0.43005508;
      R_g[10,7] := -0.20688875;
      R_g[10,8] := -0.06027012;
      R_g[10,9] := -0.64978302;
      R_g[10,10] := -3.06567740;
      R_g[10,11] := 0.07423089;
      R_g[10,12] := -0.39245805;
      R_g[10,13] := -0.47311622;
      R_g[10,14] := 0.01109051;
      R_g[10,15] := 0.29882026;
      R_g[10,16] := 0.13814223;
      R_g[10,17] := 0.20718871;
      R_g[10,18] := 0.26305798;
      R_g[10,19] := 0.67279816;
      R_g[10,20] := -0.34382215;
      R_g[10,21] := 0.54345185;
      R_g[10,22] := -0.10598019;
      R_g[10,23] := 0.08217918;
      R_g[10,24] := 0.51057720;
      R_g[10,25] := 0.12764205;
      R_g[10,26] := -0.05834693;
      R_g[10,27] := -0.33600774;
      R_g[10,28] := -0.79194522;
      R_g[10,29] := 0.23496373;
      R_g[10,30] := 0.44106248;
      R_g[10,31] := 0.30241790;
      R_g[11,0] := -0.58476233;
      R_g[11,1] := -0.14529775;
      R_g[11,2] := 0.35797024;
      R_g[11,3] := -0.98983067;
      R_g[11,4] := -0.23350208;
      R_g[11,5] := -0.01090685;
      R_g[11,6] := 0.09572268;
      R_g[11,7] := -0.34057784;
      R_g[11,8] := -0.07780220;
      R_g[11,9] := 0.66075724;
      R_g[11,10] := 0.37155905;
      R_g[11,11] := -1.91718709;
      R_g[11,12] := -0.19054978;
      R_g[11,13] := 0.00117745;
      R_g[11,14] := 0.02531583;
      R_g[11,15] := 0.54559916;
      R_g[11,16] := -0.72206557;
      R_g[11,17] := 0.41052553;
      R_g[11,18] := 0.76923150;
      R_g[11,19] := 0.42283955;
      R_g[11,20] := 0.57503432;
      R_g[11,21] := -0.45318660;
      R_g[11,22] := -0.10392044;
      R_g[11,23] := 0.00871542;
      R_g[11,24] := -0.31810006;
      R_g[11,25] := -0.22565746;
      R_g[11,26] := 0.52695656;
      R_g[11,27] := 0.10441783;
      R_g[11,28] := -0.15548979;
      R_g[11,29] := 0.46666750;
      R_g[11,30] := 0.26160634;
      R_g[11,31] := -0.11614297;
      R_g[12,0] := -0.06843481;
      R_g[12,1] := 0.19540673;
      R_g[12,2] := 0.15025875;
      R_g[12,3] := -0.17717457;
      R_g[12,4] := -0.01897787;
      R_g[12,5] := -0.12403393;
      R_g[12,6] := -0.26541382;
      R_g[12,7] := -0.08917297;
      R_g[12,8] := -0.04224596;
      R_g[12,9] := 0.11475875;
      R_g[12,10] := 0.01704736;
      R_g[12,11] := 0.10504623;
      R_g[12,12] := -4.02775335;
      R_g[12,13] := 0.01978079;
      R_g[12,14] := -0.35887444;
      R_g[12,15] := 0.27456200;
      R_g[12,16] := -0.09583630;
      R_g[12,17] := 0.32744867;
      R_g[12,18] := 0.05125649;
      R_g[12,19] := -0.07387351;
      R_g[12,20] := 0.40084934;
      R_g[12,21] := -0.33384785;
      R_g[12,22] := -0.31240118;
      R_g[12,23] := 0.02225398;
      R_g[12,24] := -0.08072241;
      R_g[12,25] := -0.00490375;
      R_g[12,26] := 0.06516396;
      R_g[12,27] := -0.25415081;
      R_g[12,28] := 0.13008058;
      R_g[12,29] := 0.11933475;
      R_g[12,30] := 0.03477714;
      R_g[12,31] := 0.03646670;
      R_g[13,0] := 0.38629496;
      R_g[13,1] := 0.07071157;
      R_g[13,2] := 0.24650244;
      R_g[13,3] := 0.18347573;
      R_g[13,4] := -0.15665166;
      R_g[13,5] := 0.05339277;
      R_g[13,6] := -0.16340585;
      R_g[13,7] := 0.01221005;
      R_g[13,8] := -0.22213434;
      R_g[13,9] := -0.72161770;
      R_g[13,10] := -0.58396721;
      R_g[13,11] := 0.29109889;
      R_g[13,12] := 0.08378197;
      R_g[13,13] := -5.32335758;
      R_g[13,14] := -0.08262666;
      R_g[13,15] := -0.33685786;
      R_g[13,16] := 0.67321271;
      R_g[13,17] := -0.30890322;
      R_g[13,18] := -0.25769258;
      R_g[13,19] := -0.51831901;
      R_g[13,20] := -0.13251379;
      R_g[13,21] := 0.68274879;
      R_g[13,22] := -0.48920557;
      R_g[13,23] := -0.14783484;
      R_g[13,24] := -0.20783210;
      R_g[13,25] := 0.22938578;
      R_g[13,26] := -0.26263767;
      R_g[13,27] := -0.11215772;
      R_g[13,28] := 0.53017223;
      R_g[13,29] := 0.11203243;
      R_g[13,30] := -0.11706309;
      R_g[13,31] := 0.81829584;
      R_g[14,0] := 0.34660137;
      R_g[14,1] := 0.30283341;
      R_g[14,2] := 0.39604405;
      R_g[14,3] := 0.34106550;
      R_g[14,4] := 0.18550380;
      R_g[14,5] := -0.15779802;
      R_g[14,6] := -0.30765054;
      R_g[14,7] := -0.05268650;
      R_g[14,8] := 0.59376097;
      R_g[14,9] := -0.12841575;
      R_g[14,10] := 0.11813307;
      R_g[14,11] := 0.16402982;
      R_g[14,12] := -0.11165220;
      R_g[14,13] := 0.09073506;
      R_g[14,14] := -1.40378904;
      R_g[14,15] := -0.07995865;
      R_g[14,16] := 0.22033221;
      R_g[14,17] := 0.23644838;
      R_g[14,18] := -0.36808783;
      R_g[14,19] := 0.37166989;
      R_g[14,20] := -0.54897916;
      R_g[14,21] := -0.46833992;
      R_g[14,22] := -0.18378656;
      R_g[14,23] := -0.48857602;
      R_g[14,24] := -0.27309927;
      R_g[14,25] := 0.23069362;
      R_g[14,26] := -0.00293107;
      R_g[14,27] := -0.25328305;
      R_g[14,28] := -0.02294313;
      R_g[14,29] := 0.34992114;
      R_g[14,30] := -0.23573494;
      R_g[14,31] := -0.23694797;
      R_g[15,0] := -0.32915220;
      R_g[15,1] := 0.17261012;
      R_g[15,2] := 0.13260838;
      R_g[15,3] := -0.39182767;
      R_g[15,4] := -0.05389502;
      R_g[15,5] := -0.11013415;
      R_g[15,6] := 0.27497944;
      R_g[15,7] := -0.14144756;
      R_g[15,8] := 0.08878060;
      R_g[15,9] := 0.07252900;
      R_g[15,10] := 0.37448993;
      R_g[15,11] := -0.36873263;
      R_g[15,12] := -0.22986236;
      R_g[15,13] := -0.34905830;
      R_g[15,14] := -0.10883336;
      R_g[15,15] := -3.20571876;
      R_g[15,16] := -0.59551466;
      R_g[15,17] := 0.36074498;
      R_g[15,18] := 0.49388149;
      R_g[15,19] := 0.17852788;
      R_g[15,20] := 0.14757296;
      R_g[15,21] := -0.23762815;
      R_g[15,22] := -0.17565729;
      R_g[15,23] := -0.13986650;
      R_g[15,24] := 0.09577942;
      R_g[15,25] := -0.13598628;
      R_g[15,26] := 0.12450486;
      R_g[15,27] := -0.13088575;
      R_g[15,28] := -0.11713267;
      R_g[15,29] := -0.03896376;
      R_g[15,30] := 0.04862077;
      R_g[15,31] := 0.15984176;
      R_g[16,0] := -0.30264369;
      R_g[16,1] := -0.32525498;
      R_g[16,2] := -0.04186732;
      R_g[16,3] := -0.23271780;
      R_g[16,4] := -0.04919057;
      R_g[16,5] := -0.07270057;
      R_g[16,6] := -0.13518807;
      R_g[16,7] := 0.21905518;
      R_g[16,8] := 0.16975564;
      R_g[16,9] := -0.27546489;
      R_g[16,10] := 0.00955923;
      R_g[16,11] := 0.23935096;
      R_g[16,12] := 0.33675262;
      R_g[16,13] := 0.04871057;
      R_g[16,14] := 0.17939901;
      R_g[16,15] := -0.05443006;
      R_g[16,16] := -1.38301742;
      R_g[16,17] := -0.62664372;
      R_g[16,18] := -0.68484670;
      R_g[16,19] := -0.24289519;
      R_g[16,20] := 0.51340222;
      R_g[16,21] := -0.10810491;
      R_g[16,22] := 0.36045137;
      R_g[16,23] := 0.25725657;
      R_g[16,24] := -0.12373380;
      R_g[16,25] := -0.48830375;
      R_g[16,26] := -0.00226057;
      R_g[16,27] := -0.17403892;
      R_g[16,28] := 0.09202776;
      R_g[16,29] := -0.20320140;
      R_g[16,30] := 0.09088694;
      R_g[16,31] := 0.03767700;
      R_g[17,0] := -0.07963943;
      R_g[17,1] := 0.01088243;
      R_g[17,2] := -0.10381653;
      R_g[17,3] := 0.40573129;
      R_g[17,4] := -0.19759901;
      R_g[17,5] := 0.13812070;
      R_g[17,6] := -0.54726249;
      R_g[17,7] := -0.34162620;
      R_g[17,8] := -0.52687168;
      R_g[17,9] := 0.15862294;
      R_g[17,10] := -0.83848864;
      R_g[17,11] := 0.30568445;
      R_g[17,12] := -0.67406219;
      R_g[17,13] := 0.53329003;
      R_g[17,14] := 0.07970227;
      R_g[17,15] := -0.48547351;
      R_g[17,16] := 0.73188645;
      R_g[17,17] := -1.73625600;
      R_g[17,18] := -0.08056269;
      R_g[17,19] := -0.54796600;
      R_g[17,20] := -0.28392172;
      R_g[17,21] := 0.52714902;
      R_g[17,22] := 0.05843952;
      R_g[17,23] := -0.00968308;
      R_g[17,24] := -0.32922518;
      R_g[17,25] := 0.13159449;
      R_g[17,26] := -0.54992115;
      R_g[17,27] := -0.05994290;
      R_g[17,28] := 0.04627676;
      R_g[17,29] := 0.11940509;
      R_g[17,30] := -0.21563587;
      R_g[17,31] := 0.49170157;
      R_g[18,0] := 0.16529544;
      R_g[18,1] := 0.14630707;
      R_g[18,2] := -0.10661374;
      R_g[18,3] := 0.31340161;
      R_g[18,4] := 0.06370668;
      R_g[18,5] := -0.17370452;
      R_g[18,6] := 0.49556559;
      R_g[18,7] := 0.43001127;
      R_g[18,8] := -0.18219198;
      R_g[18,9] := -0.46259615;
      R_g[18,10] := 0.09551673;
      R_g[18,11] := 0.46376628;
      R_g[18,12] := 0.29390970;
      R_g[18,13] := 0.54861808;
      R_g[18,14] := -0.25303873;
      R_g[18,15] := 0.01597459;
      R_g[18,16] := 0.38367042;
      R_g[18,17] := 0.25237441;
      R_g[18,18] := -1.05927384;
      R_g[18,19] := -0.53405875;
      R_g[18,20] := -0.18068475;
      R_g[18,21] := 0.21114974;
      R_g[18,22] := -0.11147468;
      R_g[18,23] := -0.10008466;
      R_g[18,24] := -0.25534129;
      R_g[18,25] := 0.36120373;
      R_g[18,26] := 0.44671911;
      R_g[18,27] := 0.12036955;
      R_g[18,28] := 0.36703530;
      R_g[18,29] := 0.06302043;
      R_g[18,30] := -0.12212825;
      R_g[18,31] := 0.30713624;
      R_g[19,0] := -0.14718637;
      R_g[19,1] := -0.08422373;
      R_g[19,2] := -0.06347395;
      R_g[19,3] := -0.52513695;
      R_g[19,4] := -0.18549855;
      R_g[19,5] := 0.07140841;
      R_g[19,6] := -0.13749593;
      R_g[19,7] := -0.12054287;
      R_g[19,8] := -0.25248626;
      R_g[19,9] := 0.51172608;
      R_g[19,10] := 0.17334092;
      R_g[19,11] := -0.56489760;
      R_g[19,12] := -0.10485484;
      R_g[19,13] := 0.16041590;
      R_g[19,14] := -0.34762689;
      R_g[19,15] := 0.32170716;
      R_g[19,16] := -0.63613361;
      R_g[19,17] := 0.45124754;
      R_g[19,18] := 0.11488474;
      R_g[19,19] := -2.78111172;
      R_g[19,20] := 0.00265766;
      R_g[19,21] := 0.19044042;
      R_g[19,22] := 0.17125109;
      R_g[19,23] := 0.05417626;
      R_g[19,24] := -0.36312413;
      R_g[19,25] := -0.21029212;
      R_g[19,26] := 0.12039141;
      R_g[19,27] := -0.21322142;
      R_g[19,28] := 0.15270446;
      R_g[19,29] := 0.18372980;
      R_g[19,30] := 0.09317994;
      R_g[19,31] := -0.11492839;
      R_g[20,0] := -0.57437384;
      R_g[20,1] := 0.40688431;
      R_g[20,2] := -0.45890683;
      R_g[20,3] := -0.19283347;
      R_g[20,4] := 0.16437508;
      R_g[20,5] := 0.01708850;
      R_g[20,6] := 0.03789070;
      R_g[20,7] := -0.21501006;
      R_g[20,8] := -0.21371005;
      R_g[20,9] := 0.51101011;
      R_g[20,10] := -0.34550032;
      R_g[20,11] := -0.50905913;
      R_g[20,12] := -0.33089176;
      R_g[20,13] := -0.57485926;
      R_g[20,14] := 0.10103830;
      R_g[20,15] := -0.69291186;
      R_g[20,16] := 0.02919241;
      R_g[20,17] := 0.52088165;
      R_g[20,18] := 0.24987195;
      R_g[20,19] := 0.33181629;
      R_g[20,20] := -4.74372387;
      R_g[20,21] := -0.27119166;
      R_g[20,22] := 0.49839181;
      R_g[20,23] := -0.19823121;
      R_g[20,24] := 0.38002643;
      R_g[20,25] := -0.42255640;
      R_g[20,26] := 0.70276517;
      R_g[20,27] := 0.40688542;
      R_g[20,28] := -0.33419290;
      R_g[20,29] := 0.00847724;
      R_g[20,30] := 0.10579581;
      R_g[20,31] := -0.28077468;
      R_g[21,0] := -0.11959543;
      R_g[21,1] := -0.37325054;
      R_g[21,2] := 0.38401762;
      R_g[21,3] := 0.36920345;
      R_g[21,4] := -0.04966644;
      R_g[21,5] := 0.13035867;
      R_g[21,6] := 0.22772673;
      R_g[21,7] := 0.12674086;
      R_g[21,8] := 0.12860185;
      R_g[21,9] := -0.91260582;
      R_g[21,10] := -0.14680338;
      R_g[21,11] := 0.23418640;
      R_g[21,12] := 0.20753485;
      R_g[21,13] := 0.55189615;
      R_g[21,14] := 0.27889958;
      R_g[21,15] := 0.29167286;
      R_g[21,16] := 0.58275050;
      R_g[21,17] := -0.86559689;
      R_g[21,18] := -0.05651870;
      R_g[21,19] := -0.29276624;
      R_g[21,20] := 0.03086585;
      R_g[21,21] := -5.40596533;
      R_g[21,22] := -0.09884489;
      R_g[21,23] := 0.17702757;
      R_g[21,24] := -0.50332761;
      R_g[21,25] := 0.41806328;
      R_g[21,26] := -0.15411623;
      R_g[21,27] := 0.41159013;
      R_g[21,28] := -0.08526843;
      R_g[21,29] := -0.07932646;
      R_g[21,30] := -0.09842971;
      R_g[21,31] := 0.33348098;
      R_g[22,0] := 0.00762757;
      R_g[22,1] := 0.07862197;
      R_g[22,2] := 0.37387678;
      R_g[22,3] := -0.49571261;
      R_g[22,4] := -0.57017809;
      R_g[22,5] := 0.00738851;
      R_g[22,6] := -0.39292586;
      R_g[22,7] := -0.16254091;
      R_g[22,8] := 0.20679110;
      R_g[22,9] := -0.12854166;
      R_g[22,10] := -0.09474767;
      R_g[22,11] := 0.21647826;
      R_g[22,12] := -0.06532618;
      R_g[22,13] := 0.35565335;
      R_g[22,14] := -0.01627116;
      R_g[22,15] := 0.66892481;
      R_g[22,16] := -0.26239413;
      R_g[22,17] := 0.05918094;
      R_g[22,18] := 0.55231690;
      R_g[22,19] := -0.35138252;
      R_g[22,20] := 0.07356476;
      R_g[22,21] := 0.07039919;
      R_g[22,22] := -1.44491446;
      R_g[22,23] := -0.21653385;
      R_g[22,24] := -0.30818766;
      R_g[22,25] := 0.26492900;
      R_g[22,26] := -0.48143271;
      R_g[22,27] := -0.45604834;
      R_g[22,28] := 0.36655438;
      R_g[22,29] := -0.29421830;
      R_g[22,30] := -0.18802145;
      R_g[22,31] := 0.22934850;
      R_g[23,0] := 0.16127868;
      R_g[23,1] := 0.03488369;
      R_g[23,2] := 0.26618156;
      R_g[23,3] := 0.24419032;
      R_g[23,4] := 0.24401736;
      R_g[23,5] := -0.08577800;
      R_g[23,6] := 0.03145451;
      R_g[23,7] := -0.06789856;
      R_g[23,8] := -0.58602816;
      R_g[23,9] := -0.12644131;
      R_g[23,10] := -0.60849923;
      R_g[23,11] := 0.34254491;
      R_g[23,12] := 0.04914726;
      R_g[23,13] := 0.07732680;
      R_g[23,14] := 0.32806584;
      R_g[23,15] := 0.17021719;
      R_g[23,16] := 0.39971253;
      R_g[23,17] := -0.44129172;
      R_g[23,18] := -0.59150064;
      R_g[23,19] := 0.34513718;
      R_g[23,20] := 0.94390410;
      R_g[23,21] := -0.69873017;
      R_g[23,22] := 0.14545058;
      R_g[23,23] := -5.33458519;
      R_g[23,24] := -0.27998123;
      R_g[23,25] := -0.68877280;
      R_g[23,26] := -0.82519758;
      R_g[23,27] := 0.21571614;
      R_g[23,28] := -0.19402163;
      R_g[23,29] := 0.89288223;
      R_g[23,30] := 0.16143902;
      R_g[23,31] := 0.60134900;
      R_g[24,0] := 0.18710028;
      R_g[24,1] := -0.15337332;
      R_g[24,2] := 0.44648594;
      R_g[24,3] := 0.04546958;
      R_g[24,4] := 0.31620455;
      R_g[24,5] := 0.22811265;
      R_g[24,6] := -0.16565078;
      R_g[24,7] := 0.19062798;
      R_g[24,8] := 0.06036144;
      R_g[24,9] := -0.53184110;
      R_g[24,10] := 0.47164744;
      R_g[24,11] := 0.14683890;
      R_g[24,12] := 0.12653536;
      R_g[24,13] := 0.66923481;
      R_g[24,14] := -0.28487730;
      R_g[24,15] := 0.86880934;
      R_g[24,16] := -0.16246760;
      R_g[24,17] := 0.11796572;
      R_g[24,18] := -0.32185227;
      R_g[24,19] := 0.14823590;
      R_g[24,20] := 0.51645494;
      R_g[24,21] := 0.13301465;
      R_g[24,22] := -0.28160232;
      R_g[24,23] := 0.19082277;
      R_g[24,24] := -5.65079260;
      R_g[24,25] := 0.02658171;
      R_g[24,26] := -0.73457789;
      R_g[24,27] := -0.54523474;
      R_g[24,28] := -0.12385467;
      R_g[24,29] := 0.09046880;
      R_g[24,30] := 0.14513928;
      R_g[24,31] := -0.45494065;
      R_g[25,0] := -0.27443600;
      R_g[25,1] := 0.03466691;
      R_g[25,2] := 0.33570170;
      R_g[25,3] := 0.11149453;
      R_g[25,4] := 0.46530443;
      R_g[25,5] := -0.11708166;
      R_g[25,6] := 0.13474351;
      R_g[25,7] := -0.01386565;
      R_g[25,8] := -0.07621623;
      R_g[25,9] := -0.65579480;
      R_g[25,10] := 0.59561032;
      R_g[25,11] := 0.70976484;
      R_g[25,12] := -0.00653760;
      R_g[25,13] := -0.11416042;
      R_g[25,14] := -0.17389505;
      R_g[25,15] := -0.29510951;
      R_g[25,16] := 0.58239830;
      R_g[25,17] := -0.31982592;
      R_g[25,18] := -0.58541101;
      R_g[25,19] := 0.11533535;
      R_g[25,20] := 0.78283572;
      R_g[25,21] := -0.67361659;
      R_g[25,22] := 0.20763648;
      R_g[25,23] := -0.07323722;
      R_g[25,24] := -0.00309061;
      R_g[25,25] := -2.58499789;
      R_g[25,26] := -0.38574260;
      R_g[25,27] := -0.09347695;
      R_g[25,28] := 0.00925173;
      R_g[25,29] := -0.02562001;
      R_g[25,30] := -0.24483223;
      R_g[25,31] := -0.02793610;
      R_g[26,0] := -0.13916478;
      R_g[26,1] := 0.08952229;
      R_g[26,2] := -0.01284268;
      R_g[26,3] := -0.16720267;
      R_g[26,4] := 0.05355829;
      R_g[26,5] := 0.00094628;
      R_g[26,6] := 0.56416976;
      R_g[26,7] := -0.17764013;
      R_g[26,8] := 0.00030415;
      R_g[26,9] := 0.37653178;
      R_g[26,10] := 0.21606593;
      R_g[26,11] := -0.31485733;
      R_g[26,12] := -0.22670522;
      R_g[26,13] := 0.12620437;
      R_g[26,14] := -0.25763687;
      R_g[26,15] := 0.28419259;
      R_g[26,16] := -0.18254681;
      R_g[26,17] := 0.37639672;
      R_g[26,18] := 0.12961774;
      R_g[26,19] := 0.13076392;
      R_g[26,20] := -0.09765223;
      R_g[26,21] := 0.05374378;
      R_g[26,22] := 0.13749219;
      R_g[26,23] := 0.02469457;
      R_g[26,24] := -0.35162118;
      R_g[26,25] := -0.18467587;
      R_g[26,26] := -3.12925005;
      R_g[26,27] := 0.19326638;
      R_g[26,28] := -0.25112805;
      R_g[26,29] := 0.16907126;
      R_g[26,30] := -0.02271179;
      R_g[26,31] := -0.16309664;
      R_g[27,0] := 0.05380776;
      R_g[27,1] := -0.15868004;
      R_g[27,2] := 0.08581222;
      R_g[27,3] := -0.02752372;
      R_g[27,4] := -0.18844807;
      R_g[27,5] := -0.02770043;
      R_g[27,6] := -0.18113151;
      R_g[27,7] := 0.21990371;
      R_g[27,8] := -0.05742185;
      R_g[27,9] := -0.04073276;
      R_g[27,10] := 0.31976753;
      R_g[27,11] := -0.10800895;
      R_g[27,12] := 0.49202874;
      R_g[27,13] := -0.11896946;
      R_g[27,14] := 0.19639397;
      R_g[27,15] := -0.16599196;
      R_g[27,16] := -0.32532701;
      R_g[27,17] := -0.03120326;
      R_g[27,18] := -0.00085085;
      R_g[27,19] := -0.04067923;
      R_g[27,20] := -0.02444752;
      R_g[27,21] := -0.06556602;
      R_g[27,22] := -0.00123137;
      R_g[27,23] := 0.02660684;
      R_g[27,24] := 0.24881741;
      R_g[27,25] := 0.04752129;
      R_g[27,26] := 0.72469455;
      R_g[27,27] := -4.37491941;
      R_g[27,28] := 0.25734231;
      R_g[27,29] := -0.47631449;
      R_g[27,30] := 0.23449393;
      R_g[27,31] := 0.31841466;
      R_g[28,0] := 0.20221227;
      R_g[28,1] := -0.19762599;
      R_g[28,2] := 0.49528366;
      R_g[28,3] := 0.60212618;
      R_g[28,4] := 0.35616049;
      R_g[28,5] := -0.29223838;
      R_g[28,6] := -0.02563414;
      R_g[28,7] := 0.25474840;
      R_g[28,8] := -0.10689805;
      R_g[28,9] := -0.53411239;
      R_g[28,10] := 0.11637564;
      R_g[28,11] := 0.50354278;
      R_g[28,12] := 0.18490633;
      R_g[28,13] := 0.10425948;
      R_g[28,14] := -0.11311629;
      R_g[28,15] := 0.17061687;
      R_g[28,16] := 0.57895732;
      R_g[28,17] := 0.44849101;
      R_g[28,18] := -0.44649935;
      R_g[28,19] := -0.08873259;
      R_g[28,20] := 0.17786060;
      R_g[28,21] := -0.34329164;
      R_g[28,22] := 0.30612892;
      R_g[28,23] := 0.32047638;
      R_g[28,24] := -0.23175892;
      R_g[28,25] := -0.06203485;
      R_g[28,26] := -0.51245290;
      R_g[28,27] := -0.07878353;
      R_g[28,28] := -2.45489097;
      R_g[28,29] := 0.29863673;
      R_g[28,30] := -0.26497275;
      R_g[28,31] := 0.39185554;
      R_g[29,0] := 0.37391195;
      R_g[29,1] := -0.06703693;
      R_g[29,2] := 0.23825873;
      R_g[29,3] := -0.37816796;
      R_g[29,4] := 0.65244371;
      R_g[29,5] := 0.01531291;
      R_g[29,6] := 0.96124893;
      R_g[29,7] := 0.05350476;
      R_g[29,8] := -0.34572360;
      R_g[29,9] := 0.67539364;
      R_g[29,10] := 0.61322534;
      R_g[29,11] := -0.22475308;
      R_g[29,12] := 0.02308607;
      R_g[29,13] := -0.10172559;
      R_g[29,14] := -0.98754531;
      R_g[29,15] := 0.27411634;
      R_g[29,16] := 0.06569140;
      R_g[29,17] := 0.97577053;
      R_g[29,18] := -0.42770064;
      R_g[29,19] := 0.51083672;
      R_g[29,20] := -0.16906519;
      R_g[29,21] := -0.55010068;
      R_g[29,22] := 0.68050390;
      R_g[29,23] := -0.01181685;
      R_g[29,24] := -0.55285066;
      R_g[29,25] := -0.37759227;
      R_g[29,26] := 0.52093881;
      R_g[29,27] := 0.36068153;
      R_g[29,28] := -0.72342020;
      R_g[29,29] := -4.50586176;
      R_g[29,30] := 0.15881208;
      R_g[29,31] := -0.55467165;
      R_g[30,0] := -0.13616283;
      R_g[30,1] := 0.11574730;
      R_g[30,2] := -0.19309571;
      R_g[30,3] := -0.11292652;
      R_g[30,4] := -0.22493608;
      R_g[30,5] := -0.09130344;
      R_g[30,6] := -0.06959558;
      R_g[30,7] := -0.08501418;
      R_g[30,8] := -0.04573239;
      R_g[30,9] := -0.44409916;
      R_g[30,10] := 0.14662819;
      R_g[30,11] := 0.11543083;
      R_g[30,12] := -0.13248284;
      R_g[30,13] := -0.12553847;
      R_g[30,14] := 0.21599039;
      R_g[30,15] := -0.11708613;
      R_g[30,16] := -0.45530063;
      R_g[30,17] := -0.03297282;
      R_g[30,18] := 0.68778771;
      R_g[30,19] := -0.25041902;
      R_g[30,20] := -0.51769501;
      R_g[30,21] := 0.72275919;
      R_g[30,22] := 0.14530140;
      R_g[30,23] := -0.10847361;
      R_g[30,24] := 0.05144800;
      R_g[30,25] := 0.34853870;
      R_g[30,26] := 0.18356445;
      R_g[30,27] := -0.50636202;
      R_g[30,28] := -0.42624116;
      R_g[30,29] := 0.33413792;
      R_g[30,30] := -2.07303715;
      R_g[30,31] := 0.24760248;
      R_g[31,0] := 0.26806670;
      R_g[31,1] := 0.04162320;
      R_g[31,2] := -0.16281062;
      R_g[31,3] := 0.30117255;
      R_g[31,4] := 0.59953493;
      R_g[31,5] := 0.02539725;
      R_g[31,6] := -0.19451533;
      R_g[31,7] := 0.02981221;
      R_g[31,8] := -0.06214313;
      R_g[31,9] := -0.37511563;
      R_g[31,10] := 0.09037945;
      R_g[31,11] := 0.34381717;
      R_g[31,12] := -0.04667491;
      R_g[31,13] := -0.22442332;
      R_g[31,14] := -0.25916281;
      R_g[31,15] := -0.52725250;
      R_g[31,16] := 0.06207185;
      R_g[31,17] := -0.30204186;
      R_g[31,18] := -0.30063924;
      R_g[31,19] := 0.24509397;
      R_g[31,20] := -0.00968230;
      R_g[31,21] := -0.19844310;
      R_g[31,22] := -0.01061517;
      R_g[31,23] := -0.21425767;
      R_g[31,24] := 0.87093484;
      R_g[31,25] := -0.09974278;
      R_g[31,26] := 0.19533432;
      R_g[31,27] := -0.09991560;
      R_g[31,28] := -0.12375148;
      R_g[31,29] := -0.20701221;
      R_g[31,30] := 0.04243100;
      R_g[31,31] := -4.28730106;
      R_o[0,0] := 0.75263089;
      R_o[0,1] := 0.03772703;
      R_o[0,2] := 0.74723381;
      R_o[0,3] := 0.04595473;
      R_o[0,4] := 1.02867210;
      R_o[0,5] := 0.40000448;
      R_o[0,6] := 0.06625949;
      R_o[0,7] := -0.08824018;
      R_o[0,8] := -0.53794587;
      R_o[0,9] := -0.52068585;
      R_o[0,10] := 0.41887417;
      R_o[0,11] := -0.98631477;
      R_o[0,12] := -0.06155511;
      R_o[0,13] := -0.61691457;
      R_o[0,14] := -0.19803670;
      R_o[0,15] := -0.30558223;
      R_o[0,16] := 0.87150252;
      R_o[0,17] := -0.18654075;
      R_o[0,18] := -0.07509329;
      R_o[0,19] := -0.33496106;
      R_o[0,20] := -0.06024283;
      R_o[0,21] := -0.04778825;
      R_o[0,22] := -0.03308541;
      R_o[0,23] := 0.54209471;
      R_o[0,24] := 0.09922121;
      R_o[0,25] := 0.00853778;
      R_o[0,26] := 0.32219675;
      R_o[0,27] := -0.13909833;
      R_o[0,28] := -0.23203412;
      R_o[0,29] := 0.00487505;
      R_o[0,30] := 0.00664908;
      R_o[0,31] := -0.21350528;
      R_o[1,0] := 0.12595357;
      R_o[1,1] := 0.56827277;
      R_o[1,2] := 0.59130812;
      R_o[1,3] := -0.17757864;
      R_o[1,4] := 0.87075138;
      R_o[1,5] := 0.20045537;
      R_o[1,6] := -0.30204454;
      R_o[1,7] := -0.05794754;
      R_o[1,8] := 1.00222409;
      R_o[1,9] := -1.44947207;
      R_o[1,10] := 0.71026599;
      R_o[1,11] := -0.64808130;
      R_o[1,12] := 0.26644772;
      R_o[1,13] := -0.07414222;
      R_o[1,14] := 1.09207368;
      R_o[1,15] := 0.68705672;
      R_o[1,16] := -0.28194490;
      R_o[1,17] := -0.35570577;
      R_o[1,18] := 0.21907447;
      R_o[1,19] := 0.08211391;
      R_o[1,20] := -0.30373713;
      R_o[1,21] := 0.01875241;
      R_o[1,22] := -0.16900432;
      R_o[1,23] := 0.19228205;
      R_o[1,24] := 0.17892483;
      R_o[1,25] := -0.21850333;
      R_o[1,26] := 0.48114797;
      R_o[1,27] := 0.11052263;
      R_o[1,28] := -0.51776105;
      R_o[1,29] := 0.89940792;
      R_o[1,30] := 1.14441526;
      R_o[1,31] := 0.04218534;
      R_o[2,0] := 0.58408523;
      R_o[2,1] := 0.68281782;
      R_o[2,2] := -3.31440473;
      R_o[2,3] := -0.29877236;
      R_o[2,4] := 1.40713286;
      R_o[2,5] := -4.67859840;
      R_o[2,6] := 1.68819666;
      R_o[2,7] := 0.25548497;
      R_o[2,8] := -0.20119862;
      R_o[2,9] := -0.69099087;
      R_o[2,10] := 0.68029040;
      R_o[2,11] := 0.07665642;
      R_o[2,12] := -0.50129002;
      R_o[2,13] := -4.08827734;
      R_o[2,14] := 0.18567920;
      R_o[2,15] := 0.45275915;
      R_o[2,16] := 0.52613461;
      R_o[2,17] := 0.75330484;
      R_o[2,18] := -0.16599981;
      R_o[2,19] := 0.79693729;
      R_o[2,20] := -0.51162231;
      R_o[2,21] := -0.81283909;
      R_o[2,22] := 0.29234949;
      R_o[2,23] := -0.28847888;
      R_o[2,24] := 4.76584196;
      R_o[2,25] := -0.15414913;
      R_o[2,26] := -0.46438026;
      R_o[2,27] := 5.13527155;
      R_o[2,28] := -0.28725153;
      R_o[2,29] := 0.26346070;
      R_o[2,30] := 0.18745001;
      R_o[2,31] := 3.02505755;
      R_o[3,0] := 0.31068292;
      R_o[3,1] := -0.22183970;
      R_o[3,2] := -0.01704333;
      R_o[3,3] := 2.34024119;
      R_o[3,4] := 1.29183245;
      R_o[3,5] := -0.06877047;
      R_o[3,6] := -0.43161812;
      R_o[3,7] := 0.16073468;
      R_o[3,8] := -0.12328651;
      R_o[3,9] := -1.27060747;
      R_o[3,10] := 0.04823594;
      R_o[3,11] := 0.29590157;
      R_o[3,12] := -0.01082665;
      R_o[3,13] := 0.33476490;
      R_o[3,14] := 0.32144535;
      R_o[3,15] := -1.52760243;
      R_o[3,16] := 0.67008370;
      R_o[3,17] := -0.15154026;
      R_o[3,18] := -1.36349714;
      R_o[3,19] := -0.27704147;
      R_o[3,20] := 0.15612660;
      R_o[3,21] := -0.06938083;
      R_o[3,22] := -0.01094813;
      R_o[3,23] := -0.04027414;
      R_o[3,24] := -0.19926009;
      R_o[3,25] := -0.06350851;
      R_o[3,26] := 0.09604281;
      R_o[3,27] := -0.42608771;
      R_o[3,28] := 0.42933077;
      R_o[3,29] := -0.12412219;
      R_o[3,30] := -0.12184074;
      R_o[3,31] := 0.30757326;
      R_o[4,0] := -0.22506563;
      R_o[4,1] := -0.00810728;
      R_o[4,2] := -0.02143744;
      R_o[4,3] := -0.34644258;
      R_o[4,4] := -0.42151707;
      R_o[4,5] := 0.25946990;
      R_o[4,6] := -0.40888065;
      R_o[4,7] := 0.36540431;
      R_o[4,8] := -0.11601024;
      R_o[4,9] := -0.06149273;
      R_o[4,10] := 0.03720159;
      R_o[4,11] := -0.32685831;
      R_o[4,12] := 0.12069022;
      R_o[4,13] := -0.46888122;
      R_o[4,14] := 0.31086460;
      R_o[4,15] := 0.14194663;
      R_o[4,16] := -0.56380451;
      R_o[4,17] := -0.50091398;
      R_o[4,18] := 0.24042240;
      R_o[4,19] := 0.34637865;
      R_o[4,20] := -0.47704268;
      R_o[4,21] := 0.33922672;
      R_o[4,22] := -0.01850082;
      R_o[4,23] := 0.18693388;
      R_o[4,24] := -0.14885549;
      R_o[4,25] := -0.15337771;
      R_o[4,26] := 0.10477851;
      R_o[4,27] := 0.03726486;
      R_o[4,28] := 0.29452741;
      R_o[4,29] := -0.19951966;
      R_o[4,30] := 0.14873424;
      R_o[4,31] := 0.33797267;
      R_o[5,0] := 0.06144769;
      R_o[5,1] := 0.40125537;
      R_o[5,2] := 0.09475308;
      R_o[5,3] := -0.19665800;
      R_o[5,4] := 0.47306305;
      R_o[5,5] := 0.88048422;
      R_o[5,6] := -0.29428431;
      R_o[5,7] := -0.02553729;
      R_o[5,8] := 0.10226711;
      R_o[5,9] := -1.00039947;
      R_o[5,10] := -0.04360576;
      R_o[5,11] := -0.92498738;
      R_o[5,12] := 0.11929558;
      R_o[5,13] := -0.20602994;
      R_o[5,14] := 0.68610996;
      R_o[5,15] := 0.22825530;
      R_o[5,16] := 0.20156530;
      R_o[5,17] := 0.32884893;
      R_o[5,18] := 0.13333681;
      R_o[5,19] := 0.33196536;
      R_o[5,20] := 0.25111938;
      R_o[5,21] := -0.51255655;
      R_o[5,22] := 0.09135021;
      R_o[5,23] := -0.11712225;
      R_o[5,24] := 0.44815740;
      R_o[5,25] := -0.30404288;
      R_o[5,26] := 0.30273652;
      R_o[5,27] := -0.10246141;
      R_o[5,28] := -0.40596756;
      R_o[5,29] := 0.21849157;
      R_o[5,30] := 0.62194777;
      R_o[5,31] := 0.34618121;
      R_o[6,0] := 0.78754842;
      R_o[6,1] := -0.53255552;
      R_o[6,2] := 0.44294843;
      R_o[6,3] := -0.62101895;
      R_o[6,4] := 0.24051274;
      R_o[6,5] := 0.08312828;
      R_o[6,6] := -0.21207847;
      R_o[6,7] := -0.63932735;
      R_o[6,8] := 0.20314510;
      R_o[6,9] := -0.56355006;
      R_o[6,10] := -0.58804530;
      R_o[6,11] := 0.70765465;
      R_o[6,12] := -0.20691018;
      R_o[6,13] := -0.28169367;
      R_o[6,14] := -0.48019099;
      R_o[6,15] := -0.12524565;
      R_o[6,16] := 0.18953465;
      R_o[6,17] := -0.59554100;
      R_o[6,18] := -0.40465477;
      R_o[6,19] := 0.35491037;
      R_o[6,20] := 0.35525450;
      R_o[6,21] := -0.79628575;
      R_o[6,22] := -0.12414181;
      R_o[6,23] := -0.13164511;
      R_o[6,24] := 0.80878896;
      R_o[6,25] := 0.23461223;
      R_o[6,26] := 0.60188603;
      R_o[6,27] := -0.60036457;
      R_o[6,28] := -0.50259900;
      R_o[6,29] := 0.64848888;
      R_o[6,30] := -0.21635155;
      R_o[6,31] := -0.37132001;
      R_o[7,0] := 0.72281468;
      R_o[7,1] := -0.36510596;
      R_o[7,2] := -0.15980141;
      R_o[7,3] := -0.49882928;
      R_o[7,4] := 0.21944484;
      R_o[7,5] := 0.33930585;
      R_o[7,6] := 0.66198981;
      R_o[7,7] := 2.29349041;
      R_o[7,8] := -1.71348310;
      R_o[7,9] := -1.17957854;
      R_o[7,10] := -0.09416397;
      R_o[7,11] := 0.17489198;
      R_o[7,12] := 0.40390244;
      R_o[7,13] := -0.37984374;
      R_o[7,14] := 0.67192376;
      R_o[7,15] := -0.60093063;
      R_o[7,16] := 0.80111188;
      R_o[7,17] := -0.14487222;
      R_o[7,18] := -0.81495136;
      R_o[7,19] := -0.57439011;
      R_o[7,20] := -0.02701034;
      R_o[7,21] := -0.21656422;
      R_o[7,22] := -0.09341363;
      R_o[7,23] := -0.40111759;
      R_o[7,24] := 1.05657363;
      R_o[7,25] := -0.05672780;
      R_o[7,26] := -0.14627363;
      R_o[7,27] := 1.03873050;
      R_o[7,28] := 0.24788009;
      R_o[7,29] := -0.26536161;
      R_o[7,30] := -0.28452447;
      R_o[7,31] := 1.08370173;
      R_o[8,0] := 0.07673319;
      R_o[8,1] := -0.68142051;
      R_o[8,2] := 0.59412581;
      R_o[8,3] := -0.32286510;
      R_o[8,4] := 0.58124644;
      R_o[8,5] := -0.54941261;
      R_o[8,6] := -0.74836421;
      R_o[8,7] := -0.08580175;
      R_o[8,8] := 0.19844094;
      R_o[8,9] := -1.80709672;
      R_o[8,10] := -0.84462225;
      R_o[8,11] := -0.72815174;
      R_o[8,12] := 0.37867835;
      R_o[8,13] := -0.09834747;
      R_o[8,14] := -0.05750175;
      R_o[8,15] := 0.24264993;
      R_o[8,16] := -0.88397968;
      R_o[8,17] := 0.84386593;
      R_o[8,18] := -0.36364627;
      R_o[8,19] := -0.46916506;
      R_o[8,20] := -0.01026842;
      R_o[8,21] := -0.22817126;
      R_o[8,22] := 0.66456556;
      R_o[8,23] := -0.20073345;
      R_o[8,24] := 0.15608832;
      R_o[8,25] := -0.33181554;
      R_o[8,26] := 0.03261386;
      R_o[8,27] := -0.17885019;
      R_o[8,28] := -1.45812154;
      R_o[8,29] := 0.46505988;
      R_o[8,30] := -0.48324671;
      R_o[8,31] := -0.35438433;
      R_o[9,0] := -0.21594478;
      R_o[9,1] := -0.20709775;
      R_o[9,2] := 0.36519870;
      R_o[9,3] := -0.73547077;
      R_o[9,4] := 0.06090719;
      R_o[9,5] := 0.16410682;
      R_o[9,6] := -0.57193118;
      R_o[9,7] := -0.07525723;
      R_o[9,8] := -0.37100428;
      R_o[9,9] := 1.03252590;
      R_o[9,10] := 0.61685145;
      R_o[9,11] := -1.23739827;
      R_o[9,12] := -0.24188256;
      R_o[9,13] := -0.11742333;
      R_o[9,14] := 0.23716070;
      R_o[9,15] := 0.02866310;
      R_o[9,16] := -0.63260299;
      R_o[9,17] := -0.02323636;
      R_o[9,18] := 0.49571911;
      R_o[9,19] := 0.80990803;
      R_o[9,20] := -0.66537541;
      R_o[9,21] := -0.83059740;
      R_o[9,22] := 0.71413642;
      R_o[9,23] := 0.39083096;
      R_o[9,24] := 0.39454761;
      R_o[9,25] := -0.75646794;
      R_o[9,26] := 0.31608939;
      R_o[9,27] := 0.16475335;
      R_o[9,28] := -0.63325989;
      R_o[9,29] := 0.68405002;
      R_o[9,30] := 0.49183965;
      R_o[9,31] := -0.64174479;
      R_o[10,0] := 0.85978961;
      R_o[10,1] := 0.38533691;
      R_o[10,2] := -0.24446277;
      R_o[10,3] := 0.43517181;
      R_o[10,4] := 0.64341557;
      R_o[10,5] := -0.37405571;
      R_o[10,6] := -0.17451185;
      R_o[10,7] := 0.39872304;
      R_o[10,8] := 0.44500470;
      R_o[10,9] := -1.23790956;
      R_o[10,10] := -2.02417660;
      R_o[10,11] := 0.06183620;
      R_o[10,12] := 0.11901627;
      R_o[10,13] := -2.94643784;
      R_o[10,14] := 0.14428562;
      R_o[10,15] := 0.27573457;
      R_o[10,16] := 0.71523923;
      R_o[10,17] := 0.06471612;
      R_o[10,18] := -0.78913754;
      R_o[10,19] := 0.15872037;
      R_o[10,20] := -0.49174178;
      R_o[10,21] := 0.18795078;
      R_o[10,22] := -0.51305294;
      R_o[10,23] := -0.13773139;
      R_o[10,24] := 3.89664268;
      R_o[10,25] := 0.79421729;
      R_o[10,26] := -0.28919408;
      R_o[10,27] := 2.04708457;
      R_o[10,28] := -0.63926643;
      R_o[10,29] := 0.00079343;
      R_o[10,30] := 0.82153952;
      R_o[10,31] := 0.78517371;
      R_o[11,0] := -0.14542149;
      R_o[11,1] := -0.05516704;
      R_o[11,2] := -0.53254628;
      R_o[11,3] := -0.12491941;
      R_o[11,4] := 1.06997979;
      R_o[11,5] := -0.07335596;
      R_o[11,6] := 0.03660922;
      R_o[11,7] := -0.62197024;
      R_o[11,8] := -0.70787662;
      R_o[11,9] := -1.29375541;
      R_o[11,10] := 1.77017760;
      R_o[11,11] := 0.15617311;
      R_o[11,12] := 0.41046301;
      R_o[11,13] := -0.07013553;
      R_o[11,14] := 0.66723573;
      R_o[11,15] := 0.58568531;
      R_o[11,16] := 0.28370255;
      R_o[11,17] := -0.72998601;
      R_o[11,18] := 0.04946580;
      R_o[11,19] := 0.05843918;
      R_o[11,20] := -0.85540062;
      R_o[11,21] := -0.97687238;
      R_o[11,22] := 0.13684957;
      R_o[11,23] := -0.55593330;
      R_o[11,24] := -0.09702116;
      R_o[11,25] := 0.66180342;
      R_o[11,26] := -0.16984765;
      R_o[11,27] := 0.12098877;
      R_o[11,28] := -0.35648933;
      R_o[11,29] := 0.39985207;
      R_o[11,30] := 0.44720337;
      R_o[11,31] := 0.31159288;
      R_o[12,0] := 0.67445350;
      R_o[12,1] := -0.62511289;
      R_o[12,2] := -0.06602924;
      R_o[12,3] := -0.07211155;
      R_o[12,4] := -0.18781437;
      R_o[12,5] := -1.00682890;
      R_o[12,6] := -0.10581888;
      R_o[12,7] := 0.65181065;
      R_o[12,8] := 0.66146719;
      R_o[12,9] := -1.83981705;
      R_o[12,10] := 0.28181201;
      R_o[12,11] := 0.36797309;
      R_o[12,12] := 2.90053463;
      R_o[12,13] := -2.21510029;
      R_o[12,14] := 1.50128496;
      R_o[12,15] := -0.82724136;
      R_o[12,16] := 1.14788032;
      R_o[12,17] := 0.03332698;
      R_o[12,18] := -0.26323086;
      R_o[12,19] := 0.50129294;
      R_o[12,20] := -0.90288156;
      R_o[12,21] := 0.31483731;
      R_o[12,22] := 1.41460466;
      R_o[12,23] := 0.37693337;
      R_o[12,24] := 0.80833459;
      R_o[12,25] := 0.69051945;
      R_o[12,26] := 0.49593949;
      R_o[12,27] := 2.64311385;
      R_o[12,28] := 0.92627031;
      R_o[12,29] := -0.26661846;
      R_o[12,30] := 0.39798808;
      R_o[12,31] := 0.27879348;
      R_o[13,0] := 0.69872397;
      R_o[13,1] := 0.09581859;
      R_o[13,2] := -0.20768847;
      R_o[13,3] := -0.28131551;
      R_o[13,4] := 0.87161541;
      R_o[13,5] := 0.17130151;
      R_o[13,6] := 0.86614621;
      R_o[13,7] := -0.73288786;
      R_o[13,8] := -0.56230539;
      R_o[13,9] := -1.29386449;
      R_o[13,10] := 0.28712273;
      R_o[13,11] := -0.38055590;
      R_o[13,12] := 0.32925129;
      R_o[13,13] := 0.11648381;
      R_o[13,14] := 0.17590009;
      R_o[13,15] := 0.47733745;
      R_o[13,16] := -0.11435314;
      R_o[13,17] := -0.25821725;
      R_o[13,18] := 0.64952123;
      R_o[13,19] := 0.43335986;
      R_o[13,20] := 0.79528856;
      R_o[13,21] := -0.31303027;
      R_o[13,22] := -0.00086104;
      R_o[13,23] := -0.60447389;
      R_o[13,24] := 2.14923382;
      R_o[13,25] := -0.30225375;
      R_o[13,26] := 0.28542003;
      R_o[13,27] := 0.20899090;
      R_o[13,28] := -0.42458954;
      R_o[13,29] := 0.82748640;
      R_o[13,30] := 0.25071397;
      R_o[13,31] := 0.33516067;
      R_o[14,0] := 0.34691715;
      R_o[14,1] := 0.44035915;
      R_o[14,2] := 0.11742699;
      R_o[14,3] := -0.25433582;
      R_o[14,4] := 0.26742107;
      R_o[14,5] := -0.02797604;
      R_o[14,6] := -0.91761684;
      R_o[14,7] := 0.00871199;
      R_o[14,8] := -0.08980305;
      R_o[14,9] := 0.00083380;
      R_o[14,10] := -0.29552653;
      R_o[14,11] := 0.17775850;
      R_o[14,12] := -0.60655963;
      R_o[14,13] := -0.65552813;
      R_o[14,14] := -1.65148222;
      R_o[14,15] := -0.03148573;
      R_o[14,16] := 0.68475866;
      R_o[14,17] := 0.48604071;
      R_o[14,18] := -0.56516480;
      R_o[14,19] := 0.04249625;
      R_o[14,20] := 0.50908113;
      R_o[14,21] := -0.94792759;
      R_o[14,22] := -0.13896449;
      R_o[14,23] := -0.58024931;
      R_o[14,24] := 0.63667297;
      R_o[14,25] := -0.18979974;
      R_o[14,26] := -0.65271628;
      R_o[14,27] := 0.36855769;
      R_o[14,28] := -0.63444155;
      R_o[14,29] := -0.16127716;
      R_o[14,30] := -0.00541620;
      R_o[14,31] := -0.32676756;
      R_o[15,0] := 0.46616146;
      R_o[15,1] := 0.13793467;
      R_o[15,2] := -1.38569939;
      R_o[15,3] := -0.21851704;
      R_o[15,4] := 2.09332156;
      R_o[15,5] := -1.44435847;
      R_o[15,6] := -0.16627391;
      R_o[15,7] := -0.29646456;
      R_o[15,8] := 4.62493992;
      R_o[15,9] := -0.73179764;
      R_o[15,10] := 0.11449970;
      R_o[15,11] := 0.32141513;
      R_o[15,12] := 0.02781674;
      R_o[15,13] := -3.39651418;
      R_o[15,14] := 0.72693330;
      R_o[15,15] := -3.30348372;
      R_o[15,16] := 0.24271241;
      R_o[15,17] := -0.69459265;
      R_o[15,18] := -0.60993481;
      R_o[15,19] := 0.50189328;
      R_o[15,20] := -2.36617303;
      R_o[15,21] := -0.73742783;
      R_o[15,22] := 1.39725518;
      R_o[15,23] := -0.17154920;
      R_o[15,24] := 4.74813509;
      R_o[15,25] := 0.86359370;
      R_o[15,26] := 0.29682380;
      R_o[15,27] := 4.01012802;
      R_o[15,28] := -0.40362200;
      R_o[15,29] := -0.32589293;
      R_o[15,30] := -0.74664325;
      R_o[15,31] := 0.69547647;
      R_o[16,0] := -0.20271565;
      R_o[16,1] := 0.28739893;
      R_o[16,2] := -0.10366275;
      R_o[16,3] := -0.63839328;
      R_o[16,4] := -0.28584042;
      R_o[16,5] := -0.21295922;
      R_o[16,6] := 0.24388939;
      R_o[16,7] := 0.04078650;
      R_o[16,8] := 0.34275502;
      R_o[16,9] := 0.40762478;
      R_o[16,10] := 0.59324360;
      R_o[16,11] := -0.53636205;
      R_o[16,12] := -0.27566653;
      R_o[16,13] := -0.23328462;
      R_o[16,14] := -0.19875692;
      R_o[16,15] := 0.22654109;
      R_o[16,16] := 0.07199147;
      R_o[16,17] := 0.44099811;
      R_o[16,18] := 0.55266190;
      R_o[16,19] := -0.17976719;
      R_o[16,20] := -0.96189427;
      R_o[16,21] := -0.15792805;
      R_o[16,22] := 0.00606035;
      R_o[16,23] := -0.51564848;
      R_o[16,24] := -0.16736200;
      R_o[16,25] := 0.10794184;
      R_o[16,26] := 0.32747260;
      R_o[16,27] := 0.52061391;
      R_o[16,28] := -0.24770921;
      R_o[16,29] := -0.11843998;
      R_o[16,30] := 0.42262232;
      R_o[16,31] := -0.67622912;
      R_o[17,0] := 1.09896290;
      R_o[17,1] := -0.64869207;
      R_o[17,2] := 0.21897116;
      R_o[17,3] := -0.34582138;
      R_o[17,4] := -1.30993581;
      R_o[17,5] := -0.05673628;
      R_o[17,6] := -1.51649237;
      R_o[17,7] := 0.00536238;
      R_o[17,8] := 0.90276903;
      R_o[17,9] := -2.21310902;
      R_o[17,10] := -0.37461346;
      R_o[17,11] := 0.83057624;
      R_o[17,12] := 0.09955819;
      R_o[17,13] := -0.79592550;
      R_o[17,14] := 0.60503864;
      R_o[17,15] := -0.56070977;
      R_o[17,16] := 0.44206971;
      R_o[17,17] := -2.85648489;
      R_o[17,18] := -0.95658404;
      R_o[17,19] := -0.66103154;
      R_o[17,20] := -0.59926432;
      R_o[17,21] := -0.11319371;
      R_o[17,22] := -1.03089595;
      R_o[17,23] := 0.16003394;
      R_o[17,24] := 3.49072146;
      R_o[17,25] := 0.41043574;
      R_o[17,26] := 0.35203537;
      R_o[17,27] := 2.91370726;
      R_o[17,28] := 0.05271170;
      R_o[17,29] := -0.20205288;
      R_o[17,30] := -0.47699225;
      R_o[17,31] := 0.73427236;
      R_o[18,0] := -0.22450200;
      R_o[18,1] := -0.07668065;
      R_o[18,2] := -0.13463168;
      R_o[18,3] := -0.79375309;
      R_o[18,4] := -0.42268148;
      R_o[18,5] := 0.16368982;
      R_o[18,6] := -0.88604885;
      R_o[18,7] := 0.18554938;
      R_o[18,8] := 0.71815532;
      R_o[18,9] := 0.25773183;
      R_o[18,10] := 0.33441162;
      R_o[18,11] := -0.26475200;
      R_o[18,12] := -0.09583112;
      R_o[18,13] := -0.33995432;
      R_o[18,14] := -0.08668236;
      R_o[18,15] := 0.53052682;
      R_o[18,16] := -0.73082268;
      R_o[18,17] := -0.00818580;
      R_o[18,18] := 0.80015409;
      R_o[18,19] := -0.38930365;
      R_o[18,20] := -0.37385350;
      R_o[18,21] := 0.26644534;
      R_o[18,22] := -0.27569091;
      R_o[18,23] := 0.16901025;
      R_o[18,24] := 0.40042493;
      R_o[18,25] := -0.76939803;
      R_o[18,26] := 0.05452700;
      R_o[18,27] := 0.09049204;
      R_o[18,28] := -0.46619353;
      R_o[18,29] := 0.74039662;
      R_o[18,30] := 0.67139417;
      R_o[18,31] := 0.11263054;
      R_o[19,0] := -0.04186005;
      R_o[19,1] := -0.02042820;
      R_o[19,2] := 0.64375228;
      R_o[19,3] := -0.98621607;
      R_o[19,4] := 1.50327301;
      R_o[19,5] := 0.91877013;
      R_o[19,6] := 0.25458473;
      R_o[19,7] := -1.09407949;
      R_o[19,8] := -0.35147515;
      R_o[19,9] := -0.75393921;
      R_o[19,10] := 0.12201059;
      R_o[19,11] := -0.15468562;
      R_o[19,12] := -0.74522096;
      R_o[19,13] := -0.95170414;
      R_o[19,14] := 0.74520445;
      R_o[19,15] := 0.34146315;
      R_o[19,16] := 0.61826760;
      R_o[19,17] := -0.19065954;
      R_o[19,18] := 0.38026699;
      R_o[19,19] := 0.97130370;
      R_o[19,20] := 0.04316740;
      R_o[19,21] := -0.41485545;
      R_o[19,22] := -0.59549576;
      R_o[19,23] := -0.17836007;
      R_o[19,24] := 0.51082230;
      R_o[19,25] := -0.13761525;
      R_o[19,26] := 0.40053996;
      R_o[19,27] := -0.79466027;
      R_o[19,28] := -0.33157697;
      R_o[19,29] := -0.58396393;
      R_o[19,30] := 0.27817172;
      R_o[19,31] := 0.54651588;
      R_o[20,0] := -0.39419258;
      R_o[20,1] := 0.27146998;
      R_o[20,2] := 0.01820673;
      R_o[20,3] := 0.29621235;
      R_o[20,4] := 0.76334292;
      R_o[20,5] := -0.65325320;
      R_o[20,6] := 0.06789777;
      R_o[20,7] := -0.40205017;
      R_o[20,8] := 0.58218980;
      R_o[20,9] := -0.69296813;
      R_o[20,10] := 0.21594040;
      R_o[20,11] := -0.35532433;
      R_o[20,12] := -0.03218510;
      R_o[20,13] := -1.00432158;
      R_o[20,14] := 0.12417480;
      R_o[20,15] := 0.92165291;
      R_o[20,16] := -0.35504830;
      R_o[20,17] := -0.28432035;
      R_o[20,18] := 0.46681264;
      R_o[20,19] := 0.88546205;
      R_o[20,20] := 0.19030854;
      R_o[20,21] := -0.58939248;
      R_o[20,22] := -0.06086200;
      R_o[20,23] := 0.12389223;
      R_o[20,24] := 1.40065300;
      R_o[20,25] := -0.38761696;
      R_o[20,26] := -0.03325392;
      R_o[20,27] := 0.04833385;
      R_o[20,28] := -0.51706809;
      R_o[20,29] := -0.84391123;
      R_o[20,30] := 0.15427513;
      R_o[20,31] := 0.02504231;
      R_o[21,0] := 0.43563822;
      R_o[21,1] := -0.05287733;
      R_o[21,2] := -0.63272291;
      R_o[21,3] := -0.38464314;
      R_o[21,4] := 0.11244948;
      R_o[21,5] := -0.34368011;
      R_o[21,6] := 0.13519558;
      R_o[21,7] := 0.17571524;
      R_o[21,8] := -0.32751995;
      R_o[21,9] := -0.54543144;
      R_o[21,10] := 0.59990895;
      R_o[21,11] := -0.33631474;
      R_o[21,12] := -0.13782535;
      R_o[21,13] := -0.65467656;
      R_o[21,14] := 0.02700578;
      R_o[21,15] := -0.33068028;
      R_o[21,16] := 0.42113748;
      R_o[21,17] := -0.49831203;
      R_o[21,18] := -0.34780854;
      R_o[21,19] := 0.11049602;
      R_o[21,20] := -0.31760716;
      R_o[21,21] := 1.28809166;
      R_o[21,22] := 0.02714989;
      R_o[21,23] := -0.14000431;
      R_o[21,24] := 2.05462027;
      R_o[21,25] := -0.04128582;
      R_o[21,26] := 0.46395308;
      R_o[21,27] := 0.14387222;
      R_o[21,28] := -0.28313118;
      R_o[21,29] := 0.21924505;
      R_o[21,30] := 0.82571280;
      R_o[21,31] := 0.77377158;
      R_o[22,0] := 0.07792897;
      R_o[22,1] := 0.20649129;
      R_o[22,2] := -0.74172878;
      R_o[22,3] := -0.58712298;
      R_o[22,4] := -0.76065350;
      R_o[22,5] := -0.46250337;
      R_o[22,6] := 0.31487158;
      R_o[22,7] := -0.74835408;
      R_o[22,8] := 1.20720458;
      R_o[22,9] := -0.62875050;
      R_o[22,10] := 0.52948600;
      R_o[22,11] := 0.02030649;
      R_o[22,12] := 0.60493541;
      R_o[22,13] := -2.44075561;
      R_o[22,14] := 0.25722051;
      R_o[22,15] := -1.02094889;
      R_o[22,16] := -0.10565599;
      R_o[22,17] := -0.10356095;
      R_o[22,18] := 0.09256380;
      R_o[22,19] := 0.93088883;
      R_o[22,20] := -1.05145490;
      R_o[22,21] := 0.07295856;
      R_o[22,22] := -0.74320340;
      R_o[22,23] := -0.80843264;
      R_o[22,24] := 1.24407017;
      R_o[22,25] := 0.27842712;
      R_o[22,26] := 0.33343524;
      R_o[22,27] := 0.36911452;
      R_o[22,28] := -0.11249841;
      R_o[22,29] := 0.74111128;
      R_o[22,30] := -0.64155215;
      R_o[22,31] := 0.55935735;
      R_o[23,0] := -0.16069618;
      R_o[23,1] := 0.58014196;
      R_o[23,2] := 0.05917757;
      R_o[23,3] := -0.36753067;
      R_o[23,4] := 0.46699741;
      R_o[23,5] := 0.07665942;
      R_o[23,6] := -0.13383338;
      R_o[23,7] := -0.06670906;
      R_o[23,8] := 0.29615077;
      R_o[23,9] := -0.18559623;
      R_o[23,10] := 0.68932790;
      R_o[23,11] := 0.13340215;
      R_o[23,12] := 0.27661046;
      R_o[23,13] := -0.44796750;
      R_o[23,14] := -0.89845961;
      R_o[23,15] := 0.08589201;
      R_o[23,16] := 0.04877722;
      R_o[23,17] := 0.59806383;
      R_o[23,18] := 0.16754775;
      R_o[23,19] := 0.08052043;
      R_o[23,20] := 0.08420350;
      R_o[23,21] := 0.05534273;
      R_o[23,22] := -0.34693667;
      R_o[23,23] := 1.55989552;
      R_o[23,24] := 0.37501606;
      R_o[23,25] := 0.10762981;
      R_o[23,26] := 0.13404730;
      R_o[23,27] := 0.00160701;
      R_o[23,28] := -0.08142579;
      R_o[23,29] := 0.68690991;
      R_o[23,30] := 0.13628589;
      R_o[23,31] := -0.29085344;
      R_o[24,0] := 0.31670842;
      R_o[24,1] := 0.78968239;
      R_o[24,2] := -0.29409191;
      R_o[24,3] := 0.46900049;
      R_o[24,4] := 0.70738745;
      R_o[24,5] := -0.13101624;
      R_o[24,6] := -0.01205759;
      R_o[24,7] := -0.38031086;
      R_o[24,8] := -0.03410443;
      R_o[24,9] := -0.43280584;
      R_o[24,10] := 0.12683180;
      R_o[24,11] := -0.50204229;
      R_o[24,12] := -0.04459752;
      R_o[24,13] := -1.82540047;
      R_o[24,14] := 0.11437972;
      R_o[24,15] := -0.25837219;
      R_o[24,16] := -0.16875745;
      R_o[24,17] := -0.30610591;
      R_o[24,18] := 0.00146165;
      R_o[24,19] := 0.57343853;
      R_o[24,20] := -0.42694604;
      R_o[24,21] := -0.32640278;
      R_o[24,22] := 0.09866292;
      R_o[24,23] := -1.04004598;
      R_o[24,24] := -0.30650541;
      R_o[24,25] := -0.44024807;
      R_o[24,26] := 1.06377351;
      R_o[24,27] := 0.15668690;
      R_o[24,28] := 0.25527728;
      R_o[24,29] := 1.11910188;
      R_o[24,30] := 0.13184597;
      R_o[24,31] := 0.66537160;
      R_o[25,0] := 0.24858460;
      R_o[25,1] := -0.21365269;
      R_o[25,2] := -0.31578684;
      R_o[25,3] := -0.23760687;
      R_o[25,4] := -0.59871852;
      R_o[25,5] := 0.04982805;
      R_o[25,6] := 0.19834036;
      R_o[25,7] := 0.12088542;
      R_o[25,8] := 0.46712711;
      R_o[25,9] := 0.63736033;
      R_o[25,10] := 0.14852153;
      R_o[25,11] := -0.34853244;
      R_o[25,12] := 0.12109412;
      R_o[25,13] := -0.52047199;
      R_o[25,14] := 0.16889386;
      R_o[25,15] := 0.26521927;
      R_o[25,16] := -0.04640898;
      R_o[25,17] := 0.14347118;
      R_o[25,18] := 0.61858296;
      R_o[25,19] := -0.65511060;
      R_o[25,20] := -0.35547650;
      R_o[25,21] := 0.10148509;
      R_o[25,22] := 0.10096559;
      R_o[25,23] := -0.28550294;
      R_o[25,24] := 0.03455871;
      R_o[25,25] := 0.67401850;
      R_o[25,26] := 0.13014895;
      R_o[25,27] := -0.28174675;
      R_o[25,28] := 0.06821958;
      R_o[25,29] := 0.32551128;
      R_o[25,30] := 0.03870281;
      R_o[25,31] := -0.16156945;
      R_o[26,0] := -0.38001239;
      R_o[26,1] := 0.56881219;
      R_o[26,2] := 0.20941640;
      R_o[26,3] := -0.48879349;
      R_o[26,4] := -0.26485169;
      R_o[26,5] := 0.05463643;
      R_o[26,6] := -0.01047605;
      R_o[26,7] := 0.06128968;
      R_o[26,8] := 0.00036229;
      R_o[26,9] := 0.59822434;
      R_o[26,10] := 0.33874771;
      R_o[26,11] := -0.82276255;
      R_o[26,12] := -0.08015160;
      R_o[26,13] := -0.24166459;
      R_o[26,14] := -0.12494149;
      R_o[26,15] := 0.25933370;
      R_o[26,16] := -0.32769927;
      R_o[26,17] := 0.58691472;
      R_o[26,18] := 0.59753895;
      R_o[26,19] := -0.06617938;
      R_o[26,20] := -0.17882954;
      R_o[26,21] := -0.17404634;
      R_o[26,22] := 0.18193702;
      R_o[26,23] := -0.03490433;
      R_o[26,24] := -0.29535082;
      R_o[26,25] := -0.03397498;
      R_o[26,26] := 0.81033039;
      R_o[26,27] := 0.03609606;
      R_o[26,28] := 0.02353646;
      R_o[26,29] := -0.01440417;
      R_o[26,30] := 0.10042611;
      R_o[26,31] := -0.04836977;
      R_o[27,0] := -0.31072620;
      R_o[27,1] := 0.44319746;
      R_o[27,2] := 0.02528284;
      R_o[27,3] := -0.15791395;
      R_o[27,4] := 0.61881942;
      R_o[27,5] := -0.03040463;
      R_o[27,6] := 0.41655910;
      R_o[27,7] := -0.73838711;
      R_o[27,8] := 0.55049175;
      R_o[27,9] := -0.43487814;
      R_o[27,10] := 0.44777703;
      R_o[27,11] := -0.00611527;
      R_o[27,12] := -0.49732092;
      R_o[27,13] := -0.21707226;
      R_o[27,14] := -0.39773074;
      R_o[27,15] := 0.64976901;
      R_o[27,16] := -0.71982020;
      R_o[27,17] := -0.01746414;
      R_o[27,18] := 0.06061571;
      R_o[27,19] := 0.38788432;
      R_o[27,20] := -0.20020573;
      R_o[27,21] := 0.41640666;
      R_o[27,22] := -0.20535807;
      R_o[27,23] := 0.30875707;
      R_o[27,24] := -0.07956075;
      R_o[27,25] := -0.12847212;
      R_o[27,26] := 0.39003900;
      R_o[27,27] := -0.80421048;
      R_o[27,28] := -0.02051540;
      R_o[27,29] := 0.11613565;
      R_o[27,30] := 0.36049625;
      R_o[27,31] := -1.31374550;
      R_o[28,0] := -0.26617476;
      R_o[28,1] := 0.63456798;
      R_o[28,2] := 0.37327421;
      R_o[28,3] := -0.50352764;
      R_o[28,4] := 0.74478012;
      R_o[28,5] := -0.59958583;
      R_o[28,6] := -0.01952661;
      R_o[28,7] := -0.27727494;
      R_o[28,8] := 0.22942626;
      R_o[28,9] := -0.18693452;
      R_o[28,10] := 0.24551098;
      R_o[28,11] := -0.18582085;
      R_o[28,12] := -0.46200407;
      R_o[28,13] := -0.33844087;
      R_o[28,14] := 0.24713075;
      R_o[28,15] := 0.41575712;
      R_o[28,16] := -0.12339561;
      R_o[28,17] := 0.63100147;
      R_o[28,18] := 0.18006700;
      R_o[28,19] := 0.59460306;
      R_o[28,20] := 0.26548737;
      R_o[28,21] := -1.45798898;
      R_o[28,22] := 0.08671085;
      R_o[28,23] := -0.13662839;
      R_o[28,24] := 0.28974804;
      R_o[28,25] := -0.36993676;
      R_o[28,26] := -0.38810381;
      R_o[28,27] := 0.18183731;
      R_o[28,28] := -0.61384946;
      R_o[28,29] := 0.88998681;
      R_o[28,30] := 0.43148291;
      R_o[28,31] := -0.01737952;
      R_o[29,0] := 0.13177893;
      R_o[29,1] := -0.05567272;
      R_o[29,2] := -2.55797052;
      R_o[29,3] := -1.07732892;
      R_o[29,4] := 1.21220803;
      R_o[29,5] := -1.56969965;
      R_o[29,6] := -2.69898748;
      R_o[29,7] := -0.28246793;
      R_o[29,8] := 0.66795498;
      R_o[29,9] := -0.37874058;
      R_o[29,10] := 0.40257087;
      R_o[29,11] := -0.41021508;
      R_o[29,12] := -0.89677757;
      R_o[29,13] := -1.41616905;
      R_o[29,14] := 0.24609458;
      R_o[29,15] := -0.72029531;
      R_o[29,16] := 0.00778214;
      R_o[29,17] := -0.71174896;
      R_o[29,18] := -0.20428607;
      R_o[29,19] := 1.29454601;
      R_o[29,20] := -0.41811258;
      R_o[29,21] := -1.16516638;
      R_o[29,22] := -0.09976852;
      R_o[29,23] := -0.60781705;
      R_o[29,24] := 1.18138075;
      R_o[29,25] := 1.49243987;
      R_o[29,26] := 0.70116144;
      R_o[29,27] := 0.88177496;
      R_o[29,28] := -0.23037660;
      R_o[29,29] := -1.76768625;
      R_o[29,30] := 0.91208470;
      R_o[29,31] := -0.19127181;
      R_o[30,0] := 0.12009788;
      R_o[30,1] := -0.06305829;
      R_o[30,2] := -0.72984314;
      R_o[30,3] := -0.38276374;
      R_o[30,4] := 0.54539680;
      R_o[30,5] := -1.35376692;
      R_o[30,6] := 0.12054427;
      R_o[30,7] := -0.11718687;
      R_o[30,8] := -0.16335595;
      R_o[30,9] := -0.39693788;
      R_o[30,10] := 1.27616143;
      R_o[30,11] := 0.38858649;
      R_o[30,12] := 0.04825598;
      R_o[30,13] := -0.69829452;
      R_o[30,14] := 0.86335611;
      R_o[30,15] := 0.25471246;
      R_o[30,16] := 0.40663683;
      R_o[30,17] := -0.13858689;
      R_o[30,18] := 0.21749221;
      R_o[30,19] := 0.72407991;
      R_o[30,20] := -0.39173615;
      R_o[30,21] := 0.05909416;
      R_o[30,22] := -0.04283657;
      R_o[30,23] := -0.93282896;
      R_o[30,24] := 1.44526589;
      R_o[30,25] := -0.16491203;
      R_o[30,26] := 0.74134064;
      R_o[30,27] := 0.47440135;
      R_o[30,28] := -0.27826020;
      R_o[30,29] := 0.86083686;
      R_o[30,30] := 2.38705564;
      R_o[30,31] := 0.59158659;
      R_o[31,0] := -0.14563540;
      R_o[31,1] := -0.46603569;
      R_o[31,2] := -0.23828754;
      R_o[31,3] := -0.21497856;
      R_o[31,4] := -0.29622266;
      R_o[31,5] := 0.07367610;
      R_o[31,6] := 0.21889332;
      R_o[31,7] := -0.23738915;
      R_o[31,8] := -0.42019483;
      R_o[31,9] := 0.39112949;
      R_o[31,10] := 0.34738326;
      R_o[31,11] := -0.50144666;
      R_o[31,12] := -0.29857567;
      R_o[31,13] := 0.08607896;
      R_o[31,14] := 0.02649515;
      R_o[31,15] := 0.56506777;
      R_o[31,16] := -0.33454859;
      R_o[31,17] := -0.10345034;
      R_o[31,18] := 0.61264884;
      R_o[31,19] := -0.31483391;
      R_o[31,20] := -0.08510064;
      R_o[31,21] := 0.76464093;
      R_o[31,22] := -0.07296492;
      R_o[31,23] := 0.38259068;
      R_o[31,24] := -0.20680594;
      R_o[31,25] := 0.07792833;
      R_o[31,26] := -0.06296873;
      R_o[31,27] := -0.13224599;
      R_o[31,28] := 0.11726132;
      R_o[31,29] := 0.27372143;
      R_o[31,30] := 0.20131113;
      R_o[31,31] := 0.34410265;
      B_i[0] := 1.05977297;
      B_i[1] := -0.77752185;
      B_i[2] := -0.05454990;
      B_i[3] := 0.88314986;
      B_i[4] := 2.16938281;
      B_i[5] := -0.58032238;
      B_i[6] := -0.70495260;
      B_i[7] := 0.20752153;
      B_i[8] := -0.44263074;
      B_i[9] := 0.39253217;
      B_i[10] := -0.80154216;
      B_i[11] := 0.79560626;
      B_i[12] := -0.00118658;
      B_i[13] := -1.62698579;
      B_i[14] := 1.40384924;
      B_i[15] := -0.13507555;
      B_i[16] := 0.55431694;
      B_i[17] := 0.71397245;
      B_i[18] := -0.00148990;
      B_i[19] := 0.21840972;
      B_i[20] := -0.27684861;
      B_i[21] := -0.80579096;
      B_i[22] := -0.24003705;
      B_i[23] := -0.58162498;
      B_i[24] := -1.42575836;
      B_i[25] := 0.38439405;
      B_i[26] := 3.43138409;
      B_i[27] := -0.96805191;
      B_i[28] := 0.30677426;
      B_i[29] := -0.86363733;
      B_i[30] := 1.65752411;
      B_i[31] := -0.05694655;
      B_f[0] := 4.11850357;
      B_f[1] := 3.80915356;
      B_f[2] := 3.32896185;
      B_f[3] := -4.06658983;
      B_f[4] := -0.78122079;
      B_f[5] := 2.33717752;
      B_f[6] := 2.97683525;
      B_f[7] := 2.31776047;
      B_f[8] := 2.21695542;
      B_f[9] := -0.30076346;
      B_f[10] := -0.82743061;
      B_f[11] := -0.74000853;
      B_f[12] := 2.29458094;
      B_f[13] := 4.44493246;
      B_f[14] := -1.22129142;
      B_f[15] := 1.71269774;
      B_f[16] := -2.14860964;
      B_f[17] := -0.00999922;
      B_f[18] := -0.01286507;
      B_f[19] := -0.24900147;
      B_f[20] := 2.74852705;
      B_f[21] := 2.75391650;
      B_f[22] := -0.26369506;
      B_f[23] := 3.12250614;
      B_f[24] := 3.50876307;
      B_f[25] := 1.24471641;
      B_f[26] := 2.86891937;
      B_f[27] := 1.47885728;
      B_f[28] := -0.03386326;
      B_f[29] := 2.28063703;
      B_f[30] := 0.76983297;
      B_f[31] := 2.23378706;
      B_g[0] := 0.67241311;
      B_g[1] := -0.63885009;
      B_g[2] := -0.90349925;
      B_g[3] := -2.79336119;
      B_g[4] := 1.65765214;
      B_g[5] := -0.83395064;
      B_g[6] := -0.21865635;
      B_g[7] := 0.23917481;
      B_g[8] := 0.29897273;
      B_g[9] := -1.96458340;
      B_g[10] := 1.01046002;
      B_g[11] := 1.69552255;
      B_g[12] := 0.52112406;
      B_g[13] := -1.21443260;
      B_g[14] := 0.42707205;
      B_g[15] := 0.30916595;
      B_g[16] := -0.51244986;
      B_g[17] := -0.99837846;
      B_g[18] := -1.55904579;
      B_g[19] := 0.59441733;
      B_g[20] := 0.25117961;
      B_g[21] := -0.76235783;
      B_g[22] := 0.18406813;
      B_g[23] := -0.52563477;
      B_g[24] := 1.11005735;
      B_g[25] := -0.20509416;
      B_g[26] := 0.40615445;
      B_g[27] := 0.81266654;
      B_g[28] := -0.99892116;
      B_g[29] := 0.04178268;
      B_g[30] := 0.42290145;
      B_g[31] := 0.12953959;
      B_o[0] := 2.36205053;
      B_o[1] := 4.44841862;
      B_o[2] := 3.44511604;
      B_o[3] := -0.27658543;
      B_o[4] := 0.62766176;
      B_o[5] := 3.89909387;
      B_o[6] := 2.23212004;
      B_o[7] := 3.08706617;
      B_o[8] := 3.04965401;
      B_o[9] := 2.26128387;
      B_o[10] := 2.17441511;
      B_o[11] := 3.20681429;
      B_o[12] := 3.75658846;
      B_o[13] := 3.67272520;
      B_o[14] := 2.05645180;
      B_o[15] := 2.52790165;
      B_o[16] := 1.83170414;
      B_o[17] := 3.62001419;
      B_o[18] := 4.37526703;
      B_o[19] := 3.76178741;
      B_o[20] := 3.90018415;
      B_o[21] := 2.82298088;
      B_o[22] := 2.73789883;
      B_o[23] := 2.35665083;
      B_o[24] := 3.36428308;
      B_o[25] := 1.81089711;
      B_o[26] := 0.79725283;
      B_o[27] := 2.29590178;
      B_o[28] := 3.59097409;
      B_o[29] := 2.43540621;
      B_o[30] := 2.37923050;
      B_o[31] := 1.37423539;
      FC_W[0,0] := -0.34967208;
      FC_W[0,1] := 0.17095216;
      FC_W[0,2] := 0.18948522;
      FC_W[0,3] := 0.43564883;
      FC_W[0,4] := -0.72084081;
      FC_W[0,5] := 0.20435235;
      FC_W[0,6] := 0.43418887;
      FC_W[0,7] := 1.39729345;
      FC_W[0,8] := -0.87131464;
      FC_W[0,9] := -0.67471236;
      FC_W[0,10] := 0.22794832;
      FC_W[0,11] := 0.14453813;
      FC_W[0,12] := -1.05575025;
      FC_W[0,13] := 0.05739802;
      FC_W[0,14] := 0.15091233;
      FC_W[0,15] := 0.88983119;
      FC_W[0,16] := -0.43641257;
      FC_W[0,17] := 0.17820166;
      FC_W[0,18] := -0.79069114;
      FC_W[0,19] := -0.23154163;
      FC_W[0,20] := 0.19985847;
      FC_W[0,21] := -0.40778121;
      FC_W[0,22] := 0.14641519;
      FC_W[0,23] := -0.24937966;
      FC_W[0,24] := 0.09585419;
      FC_W[0,25] := -0.13808215;
      FC_W[0,26] := -0.20577344;
      FC_W[0,27] := -0.17500097;
      FC_W[0,28] := 0.46872810;
      FC_W[0,29] := 0.13711151;
      FC_W[0,30] := 0.11427750;
      FC_W[0,31] := 0.82231474;
      FC_W[1,0] := 0.03423055;
      FC_W[1,1] := 0.39694929;
      FC_W[1,2] := -1.06318247;
      FC_W[1,3] := -0.16354848;
      FC_W[1,4] := 0.18805455;
      FC_W[1,5] := 0.75300908;
      FC_W[1,6] := -0.74681133;
      FC_W[1,7] := 0.60798770;
      FC_W[1,8] := 0.94372779;
      FC_W[1,9] := 0.35550115;
      FC_W[1,10] := -0.57321185;
      FC_W[1,11] := 0.33739200;
      FC_W[1,12] := 0.03249437;
      FC_W[1,13] := -0.57342994;
